      | #   log_info("Trying to find object by color:", to_str(material))
      | #   while (i < OBJECT_MAP.length()):
      | #       if (OBJECT_MAP[i].material == material):
      | #           log_info("Object model found:", to_str(OBJECT_MAP[i]))
      | #           return OBJECT_MAP[i]
      | #       end
      | #       i = i + 1
      | #   end
      | #   return OBJ_DEFAULT  # Return default pattern if not found
      | # end
      | 
      | def find_object_by_objectname(objectname):
      |     local i = 0
      |     #log_info("Trying to find object by color:", to_str(objectname))
      |     while (i < OBJECT_MAP.length()):
      |         if (OBJECT_MAP[i].obj_name == objectname):
      |             log_info("Object Model found: [" + to_str(OBJECT_MAP[i].description) + "]")
      |             return OBJECT_MAP[i]
      |         end
      |         i = i + 1
      |     end
      |     log_warning("no Object Model found for objectname:[" + to_str(objectname) + "]")
      |     return create_object()
      | end
      | 
      | def find_smallest_object():
      |     local i = 0
      |     local min_size = OBJECT_MAP[0].height
      |     #log_info("Trying to find object by color:", to_str(objectname))
      |     while (i < OBJECT_MAP.length()):
      |         if (OBJECT_MAP[i].height <= min_size and OBJECT_MAP[i].height != 0):
      |             log_info("smaller object found: [" + to_str(OBJECT_MAP[i].description) + "]")
      |             min_size = OBJECT_MAP[i].height
      |         end
      |         i = i + 1
      |     end
      |     return min_size
      | end
      | 
      | def find_gripper_config_by_objectname(objectname):
      | local i = 0
      | while (i < GRIPPER_CONFIG_MAP.length()):
      |     #log_info("gripper config:",to_str(GRIPPER_CONFIG_MAP[i]))
      |     if (GRIPPER_CONFIG_MAP[i].object == objectname):
      |         log_info("found gripper parameters [" + to_str(GRIPPER_CONFIG_MAP[i]) + "]")
      |         return GRIPPER_CONFIG_MAP[i]
      |     end
      |     i = i + 1
      | end
      | 
      | log_warning("no gripper parameters found for object type: " + to_str(objectname))
      | return create_gripper_config()
      | end
      | # Function to find a landmark by item
      | def find_landmark_by_id(lm_id):
      |     local i = 0
      |     while i < LANDMARK_MAP.length():
      |         if LANDMARK_MAP[i].lm_id == lm_id:
      |             log_info("found landmark with id(" + to_str(lm_id) + "): [" + to_str(LANDMARK_MAP[i].description) + "]")
      |             return LANDMARK_MAP[i]
      |         end
      |         i = i + 1
      |     end
      |     log_warning("landmark not found for lm_id [" + to_str(lm_id) + "]")
      |     return create_landmark()
      | end
      | # Function to find a landmark by item
      | def find_landmark_by_capture_pos(capture_pos):
      |     local i = 0
      |     while i < LANDMARK_MAP.length():
      |         if LANDMARK_MAP[i].capture_pos == capture_pos:
      |             log_info("found landmark by capture_pos [" + to_str(LANDMARK_MAP[i].description) + "]")
      |             return LANDMARK_MAP[i]
      |         end
      |         i = i + 1
      |     end
      |     log_warning("Landmark not found for capture_pos: [" + to_str(capture_pos) + "]")
      |     return create_landmark()
      | end
      | 
      | def update_landmark_by_capture_pos(capture_pos, lm_pos):
      |     local i = 0
      |     while i < LANDMARK_MAP.length():
      |         if LANDMARK_MAP[i].capture_pos == capture_pos:
      |             log_info("updated landmark from [" + to_str(LANDMARK_MAP[i].description) + "]")
      |             LANDMARK_MAP[i].actual_frame = lm_pos
      |             return True
      |         end
      |         i = i + 1
      |     end
      |     log_warning("Landmark not found for capture_pos: [" + to_str(capture_pos) + "]")
      |     return False
      | end
      | 
      | def update_landmark_by_id(lm_id,lm_pos):
      |     local i = 0
      |     while i < LANDMARK_MAP.length():
      |         if LANDMARK_MAP[i].lm_id == lm_id:
      |             log_info("updated landmark.actual_frame from [" + to_str(LANDMARK_MAP[i].description + "]"))
      |             LANDMARK_MAP[i].actual_frame = lm_pos
      |             return True
      |         end
      |         i = i + 1
      |     end
      |     log_warning("Landmark not found for lm_id " + to_str(lm_id))
      |     return False
      | end
      | 
      | def find_vision_config_by_frame(frame):
      |     local i = 0
      |     while i < VISION_CONFIG_MAP.length():
      |         if VISION_CONFIG_MAP[i].capture_pos == frame:
      |             log_info("Vision Config found: [" + to_str(VISION_CONFIG_MAP[i].description) + "]")
      |             return VISION_CONFIG_MAP[i]
      |         end
      |         i = i + 1
      |     end
      |     log_info("Vision Config not found for frame: " + to_str(frame))
      |     return create_vision_config()
      | end
      | 
      | def find_vision_config_by_itemid(id):
      |     local i = 0
      |     while i < VISION_CONFIG_MAP.length():
      |         if VISION_CONFIG_MAP[i].item_id == id:
      |             log_info("Vision Config found: [" + to_str(VISION_CONFIG_MAP[i].description) + "]")
      |             return VISION_CONFIG_MAP[i]
      |         end
      |         i = i + 1
      |     end
      |     log_info("Vision Config not found for item: " + to_str(id))
      |     return create_vision_config()
      | end
      | 
      | def find_inspect_config_by_itemid(id):
      |     local i = 0
      |     while i < INSPECT_CONFIG_MAP.length():
      |         if INSPECT_CONFIG_MAP[i].item_id == id:
      |             log_info("Inspect Config found: [" + to_str(INSPECT_CONFIG_MAP[i].description) + "]")
      |             return INSPECT_CONFIG_MAP[i]
      |         end
      |         i = i + 1
      |     end
      |     log_info("Inspect Config not found for item: " + to_str(id))
      |     return create_inspect_config()
      | end
    Script file /programs/04 Scripts/SCRIPT Device Robotiq Greifer v0.2.script
      | # ############ SCRIPT Device Robotiq Greifer ###############
      | # **********************************************************
      | # Customer          :   URG
      | # Product Name      :   uLabMobile
      | # **********************************************************
      | # Controller/Robot  :   UR5e
      | # Software          :   5.17
      | # Dependencies      :   Logs Script, Robotiq Gripper and Gripper Datastructure for args (Factory Script), URCAP Robotiq
      | # **********************************************************
      | # Author            :   D.Kreugel, P.Köhnke
      | # Copyright (c)     :   United Robotics Group Health and Food GmbH
      | #                       An der Riede 2
      | #                       28816 Stuhr
      | #                       Germany
      | # *********************************************************
      | # Description       :   Gripper Robotiq Device Interface for Robotiq E-Hand Gripper
      | # Version           :   0.2
      | # Created           :   18.07.2024
      | # Updated           :
      | # *********************************************************
      | # Modifications     :
      | #
      | # Date              :
      | # Name              :
      | # Reason            :
      | # *********************************************************
      | # TODO              :   documentation
      | 
      | # RobotiQ Gripper
      | ROBOTIQ_GRP_CLOSE = 0
      | ROBOTIQ_GRP_OPEN = 40
      | 
      | # #############FORCEMODE###############
      | ROBOTIQ_GRP_FORCE = struct(FULL=100, HALF=50, LOW=25, NONE=0)
      | 
      | # #############SPEED###################
      | ROBOTIQ_GRP_SPEED = struct(FAST=100, MEDIUM=50, SLOW=20)
      | 
      | # ############VALIDATION###############
      | ROBOTIQ_GRP_VALIDATION = struct(ON=1, OFF=0, SKIP=-1)
      | 
      | # struct(prepick=0, pick=0, place=0, force=0, speed=0, validation=0, object_type=0, description="default")
      | def gripper_robotiq_activate():
      |     return rq_activate_and_wait()
      | end
      | 
      | def gripper_robotiq_reset_and_activate():
      |     return rq_reset_and_activate()
      |     #return rq_reset()
      | end
      | 
      | def gripper_robotiq_is_activated():
      |     return rq_is_gripper_activated()
      | end
      | 
      | def gripper_robotiq_get_current_pos_mm():
      |     return rq_current_pos_mm()
      | end
      | # Function to check if the RobotiQ gripper has an object
      | def gripper_robotiq_has_object():
      |     result = rq_is_object_detected()
      |     if result == False:
      |         log_error("No object detected by the gripper")
      |     end
      |     return result
      | end
      | 
      | def gripper_robotiq_move_to_mm(mm):
      |     if(gripper_robotiq_is_activated() == False):
      |         gripper_robotiq_activate()
      |     end
      |     return rq_move_and_wait_mm(mm)
      | end
      | 
      | def gripper_robotiq_close():
      |     if(gripper_robotiq_is_activated() == False):
      |         gripper_robotiq_activate()
      |     end
      |     return rq_close_and_wait()
      | end
      | 
      | def gripper_robotiq_open():
      |     if(gripper_robotiq_is_activated() == False):
      |         gripper_robotiq_activate()
      |     end
      |     return rq_open_and_wait()
      | end
      | 
      | def gripper_robotiq_set_force(force):
      |     return rq_set_force_norm(force)
      | end
      | 
      | def gripper_robotiq_set_speed(velocity):
      |     return rq_set_speed_norm(velocity)
      | end
      | # Function to initialize the RobotiQ gripper
      | # args = struct(obj_type = object.obj_type, force = force, speed = speed, validation = validation, width = (prepick=2, pick=0, place=2))
      | def gripper_robotiq_init(args):
      |     log_info("args:"+to_str(args))
      |     gripper_robotiq_set_force(args.force)
      |     gripper_robotiq_set_speed(args.speed)
      |     if(gripper_robotiq_is_activated() == False):
      |         gripper_robotiq_activate()
      |     end
      |     log_info("Robotiq Gripper Initialized with arguments:" + to_str(args))
      |     return True
      | end
      | # Function to prepare the RobotiQ gripper for picking
      | # args = struct(obj_type = object.obj_type, force = force, speed = speed, validation = validation, width = (prepick=2, pick=0, place=2))
      | def gripper_robotiq_prepick(args):
      |     gripper_robotiq_init(args)
      | 
      |     if(args.width.prepick <= ROBOTIQ_GRP_CLOSE):
      |         rq_close_and_wait()
      |     elif(args.width.prepick >= ROBOTIQ_GRP_OPEN):
      |         rq_open_and_wait()
      |     else:
      |         rq_move_and_wait_mm(args.width.prepick)
      |     end
      | 
      |     log_info("Robotiq Gripper prepick with arguments:" + to_str(args))
      |     return True
      | end
      | 
      | # Function to place an object using the RobotiQ gripper
      | # args = struct(obj_type = object.obj_type, force = force, speed = speed, validation = validation, width = (prepick=2, pick=0, place=2))
      | def gripper_robotiq_place(args):
      |     gripper_robotiq_init(args)
      | 
      |     if(args.width.place <= ROBOTIQ_GRP_CLOSE):
      |         rq_close_and_wait()
      |     elif(args.width.place >= ROBOTIQ_GRP_OPEN):
      |         rq_open_and_wait()
      |     else:
      |         rq_move_and_wait_mm(args.width.place)
      |     end
      | 
      |     log_info("Gripper Place with arguments:"+ to_str(args))
      |     return True
      | end
      | 
      | # Function to pick an object using the RobotiQ gripper
      | # args = struct(obj_type = object.obj_type, force = force, speed = speed, validation = validation, width = (prepick=2, pick=0, place=2))
      | def gripper_robotiq_pick(args):
      |     gripper_robotiq_init(args)
      | 
      |     if(args.width.pick <= ROBOTIQ_GRP_CLOSE):
      |         rq_close_and_wait()
      |     elif(args.width.pick >= ROBOTIQ_GRP_OPEN):
      |         rq_open_and_wait()
      |     else:
      |         rq_move_and_wait_mm(args.width.pick)
      |     end
      | 
      |     log_info("Gripper Pick with arguments:" + to_str(args))
      | 
      |     if args.validation == ROBOTIQ_GRP_VALIDATION.ON:
      |         if gripper_robotiq_has_object() == False:
      |             log_error("Validation failed, no object detected")
      |             return False
      |         end
      |     end
      | 
      |     return True
      | end
      | 
      | 
      | # def gripper_robotiq_close_and_validate():
      | #     rq_close_and_wait()
      | #     if gripper_robotiq_has_object() == False:
      | #         log_error("Validation failed, no object detected")
      | #         return False
      | #     else:
      | #         return True
      | #     end
      | # end
    Script file /programs/04 Scripts/SCRIPT uLM Gripperconfig v0.6.script
      | ############# SCRIPT uLM Gripperconfig ###############
      | #*****************************************************
      | # Customer          :   URG
      | # Product Name      :   uLabMobile
      | #****************************************************
      | # Controller/Robot  :   UR5e
      | # Software          :   UR-Script
      | # Dependencies      :   physical Gripper and Datastructure from Factory for args -> Device Script and Implementations of the Functions
      | # How To            :   Assign all Functioncalls to the equivalent of the used Device Script
      | #****************************************************
      | # Author            :   D.Kreugel, P.Köhnke
      | # Copyright (c)     :   United Robotics Group Health and Food GmbH
      | #                       An der Riede 2
      | #                       28816 Stuhr
      | #                       Germany
      | #****************************************************
      | # Description       :   Defines all Gripperm related Parameters and Functions
      | # Version           :   0.6
      | # Created           :   18.07.2024
      | # Updated           :
      | #****************************************************
      | # Modifications     :   -> at the moment Gripperconfig linked to Robotiq Gripper Device Script
      | # Date              :   18.07.2017
      | # Name              :   D.Kreugel
      | # Reason            :   uLM Standard
      | #****************************************************
      | # TO DO             : Implement Activate and Reset Routine at the beginning or after an error depending on the state if an Object is gripped or not, documentation
      | 
      | 
      | 
      | # GRIPPER DEFINES
      | GRIPPER_CLOSE = ROBOTIQ_GRP_CLOSE
      | GRIPPER_OPEN = ROBOTIQ_GRP_OPEN
      | # #############FORCE###############
      | GRIPPER_FORCE = ROBOTIQ_GRP_FORCE
      | # #############SPEED###################
      | GRIPPER_SPEED = ROBOTIQ_GRP_SPEED
      | # ############VALIDATION###############
      | GRIPPER_VALIDATION = ROBOTIQ_GRP_VALIDATION
      | 
      | # takes force in %
      | def gripper_set_force(force):
      |     return gripper_robotiq_set_force(force)
      | end
      | 
      | # takes speed in %
      | def gripper_set_speed(velocity):
      |     return gripper_robotiq_set_speed(velocity)
      | end
      | 
      | def gripper_activate():
      |     return gripper_robotiq_activate()
      | end
      | 
      | def gripper_reset_and_activate():
      |     return gripper_robotiq_reset_and_activate()
      | end
      | 
      | def gripper_is_activated():
      |     return gripper_robotiq_is_activated()
      | end
      | 
      | def gripper_get_current_pos_mm():
      |     return gripper_robotiq_get_current_pos_mm()
      | end
      | 
      | def gripper_has_object():
      |     return gripper_robotiq_has_object()
      | end
      | 
      | def gripper_open():
      |     return gripper_robotiq_open()
      | end
      | 
      | def gripper_close():
      |     return gripper_robotiq_close()
      | end
      | 
      | def gripper_move_to_pos_mm(mm):
      |     return gripper_robotiq_move_to_mm(mm)
      | end
      | 
      | # args = struct(obj_type = object.obj_type, force = force, speed = speed, validation = validation, width = (prepick=2, pick=0, place=2))
      | def gripper_init(args):
      |     return gripper_robotiq_init(args)
      | end
      | 
      | # args = struct(obj_type = object.obj_type, force = force, speed = speed, validation = validation, width = (prepick=2, pick=0, place=2))
      | def gripper_prepick(args):
      |     return gripper_robotiq_prepick(args)
      | end
      | 
      | # args = struct(obj_type = object.obj_type, force = force, speed = speed, validation = validation, width = (prepick=2, pick=0, place=2))
      | def gripper_pick(args):
      |     return gripper_robotiq_pick(args)
      | end
      | 
      | # args = struct(obj_type = object.obj_type, force = force, speed = speed, validation = validation, width = (prepick=2, pick=0, place=2))
      | def gripper_place(args):
      |     return gripper_robotiq_place(args)
      | end
      | 
      | 
      | # def gripper_close_and_validate():
      | #     return gripper_robotiq_close_and_validate()
      | # end
    Script file /programs/04 Scripts/SCRIPT uLM Projectconfig 0.2.script
      | ############# SCRIPT uLM Projectconfig ###############
      | #*****************************************************
      | # Customer          :   URG
      | # Product Name      :   uLabMobile
      | #****************************************************
      | # Controller/Robot  :   UR5e
      | # Software          :   5.17
      | # Dependencies      :   Factory Script, Defines Script, relevant project knowledge about objects, patterns, items, commands, vision skills, landmarktypes and movements
      | # How To            :   Define Step by Step all Project Data by creating the objects and appending them to the assigned List, if you skip information
      | #                       the default value will be assigned -> give as many details as possible as the default values will not work in some cases
      | #****************************************************
      | # Author            :   D.Kreugel
      | # Copyright (c)     :   United Robotics Group Health and Food GmbH
      | #                       An der Riede 2
      | #                       28816 Stuhr
      | #                       Germany
      | #****************************************************
      | # Description       :   Project Related Configurations -> in the future will be configured by UGO
      | # Version           :   0.2
      | # Created           :   18.07.2024
      | # Updated           :
      | #****************************************************
      | # Modifications     :
      | # Date              :
      | # Name              :
      | # Reason            :
      | #****************************************************
      | # TO DO             :  Simplify Rack Assignment, create Enums for Choices that can be made and will be repeated in many projects, documentation
      | 
      | #
      | 
      | # Please Import DeviceScripts and Defines Script First as you may wanna use some of the Defined Variables here
      | 
      | # Define here the Objects that should be handled, add a new Object Type in the defines if necessary
      | # create_object(id=0, obj_name=0, height=0, width=0, color="default", material="default", description="default")
      | # struct(NONE=0, CC_SAMPLE=1, CC_RACK=2, COAG_SAMPLE=3, COAG_RACK=4, HEMA_SAMPLE=5, HEMA_RACK=6, INPUT_RACK=7, CF_RACK=8, ANY_SAMPLE=9, ANY_RACK=10)
      | #create_object(id=0, obj_name=0, height=0, width=0, obj_type = 0, description="default")
      | OBJECT_MAP.append(create_object(id=0, obj_name=Objects.NONE, obj_type=ObjectType.NONE, height=0, width=0, description="None Object"))
      | OBJECT_MAP.append(create_object(id=1, obj_name=Objects.CC_SAMPLE, obj_type=ObjectType.SAMPLE, height=108, width=15, description="BD Li-Heparin"))
      | OBJECT_MAP.append(create_object(id=2, obj_name=Objects.HEMA_SAMPLE, obj_type=ObjectType.SAMPLE, height=81, width=13, description="BD EDTA"))
      | OBJECT_MAP.append(create_object(id=3, obj_name=Objects.CC_SAMPLE, obj_type=ObjectType.SAMPLE, height=108, width=15, description="BD Li-Heparin"))
      | OBJECT_MAP.append(create_object(id=4, obj_name=Objects.HEMA_SAMPLE, obj_type=ObjectType.SAMPLE, height=81, width=13, description="Sarstedt EDTA"))
      | OBJECT_MAP.append(create_object(id=5, obj_name=Objects.CC_SAMPLE, obj_type=ObjectType.SAMPLE, height=110, width=15, description="Sarstedt Serum-Gel"))
      | OBJECT_MAP.append(create_object(id=6, obj_name=Objects.ANY_SAMPLE, obj_type=ObjectType.SAMPLE, height=110, width=15, description="Any Sample"))
      | OBJECT_MAP.append(create_object(id=7, obj_name=Objects.ANY_RACK, height=150, width=120, description="Any Rack"))
      | OBJECT_MAP.append(create_object(id=8, obj_name=Objects.CF_RACK, height=110, width=15, description="Centrifuge Rack"))
      | OBJECT_MAP.append(create_object(id=12, obj_name=Objects.COBAS_RACK, height=OBJECT_REFERENCE_HEIGHT, width=20, description="Cobas Rack"))
      | OBJECT_MAP.append(create_object(id=9, obj_name=Objects.TARA_SAMPLE, obj_type=ObjectType.SAMPLE, height=110, width=15, description="Tara Sample"))
      | OBJECT_MAP.append(create_object(id=10, obj_name=Objects.BUTTON, obj_type=ObjectType.BUTTON, height=0, width=0, description="Button"))
      | OBJECT_MAP.append(create_object(id=11, obj_name=Objects.XN550_DRAWER, height=OBJECT_REFERENCE_HEIGHT, width=25, description="XN550 Drawer"))
      | 
      | #create_sample(obj_id=0, diameter=0, color="", material="", description="")
      | SAMPLES = make_list(0,create_sample(),MAX_ITEM_OBJ)
      | SAMPLES.append(create_sample(obj_id=1, cap_diameter=17.4, raw_diameter=15.3, color="darkgreen", material="88", description="BD Li-Heparin -> decapped in Cobas"))
      | SAMPLES.append(create_sample(obj_id=1, cap_diameter=17.4, raw_diameter=15.3, color="darkgreen", material="80", description="BD Li-Heparin -> decapped in Cobas"))
      | SAMPLES.append(create_sample(obj_id=1, cap_diameter=17.4, raw_diameter=15.3, color="darkgreen", material="93", description="BD Li-Heparin -> decapped in archive"))
      | SAMPLES.append(create_sample(obj_id=2, cap_diameter=15.5, raw_diameter=12.3, color="violet", material="82", description="BD EDTA -> Sysmex ->Archive"))
      | SAMPLES.append(create_sample(obj_id=2, cap_diameter=15.5, raw_diameter=12.3, color="violet", material="91", description="BD EDTA ->Archive"))
      | SAMPLES.append(create_sample(obj_id=2, cap_diameter=15.5, raw_diameter=12.3, color="violet", material="96", description="BD EDTA ->Archive"))
      | SAMPLES.append(create_sample(obj_id=3, cap_diameter=17.4, raw_diameter=15.3, color="lightgreen", material="88", description="BD Li-Heparin -> decapped in Cobas"))
      | SAMPLES.append(create_sample(obj_id=3, cap_diameter=17.4, raw_diameter=15.3, color="lightgreen", material="93", description="BD Li-Heparin -> decapped in Archive"))
      | SAMPLES.append(create_sample(obj_id=3, cap_diameter=17.4, raw_diameter=15.3, color="lightgreen", material="97", description="BD Li-Heparin -> decapped in Archive"))
      | SAMPLES.append(create_sample(obj_id=4, cap_diameter=15.6, raw_diameter=12.3, color="red", material="82", description="BD EDTA -> Sysmex ->Archive"))
      | SAMPLES.append(create_sample(obj_id=4, cap_diameter=15.6, raw_diameter=12.3, color="red", material="91", description="BD EDTA -> Archive"))
      | SAMPLES.append(create_sample(obj_id=4, cap_diameter=15.6, raw_diameter=12.3, color="red", material="96", description="BD EDTA -> Archive"))
      | SAMPLES.append(create_sample(obj_id=5, cap_diameter=17.4, raw_diameter=15.3, color="brown", material="80", description="Sarstedt Serum-Gel -> decapped in Cobas"))
      | SAMPLES.append(create_sample(obj_id=5, cap_diameter=17.4, raw_diameter=15.3, color="brown", material="93", description="Sarstedt Serum-Gel -> decapped in Archive"))
      | 
      | # Gripper Configurations depending on the Object Type , add new force and speed in the Defines if necessary
      | # create_gripper_config(gripper_offset=struct(prepick=2, pick=0, place=2), force=0, speed=0, validation=0, object=create_object())
      | GRIPPER_CONFIG_MAP.append(create_gripper_config(gripper_offset=struct(prepick=2, pick=0, place=2), force=GRIPPER_FORCE.HALF, speed=GRIPPER_SPEED.MEDIUM, validation=GRIPPER_VALIDATION.ON, object=find_object_by_objectname(Objects.ANY_SAMPLE)))
      | GRIPPER_CONFIG_MAP.append(create_gripper_config(gripper_offset=struct(prepick=2, pick=0, place=2), force=GRIPPER_FORCE.FULL, speed=GRIPPER_SPEED.MEDIUM, validation=GRIPPER_VALIDATION.ON, object=find_object_by_objectname(Objects.ANY_RACK)))
      | GRIPPER_CONFIG_MAP.append(create_gripper_config(gripper_offset=struct(prepick=2, pick=0, place=2), force=GRIPPER_FORCE.HALF, speed=GRIPPER_SPEED.MEDIUM, validation=GRIPPER_VALIDATION.ON, object=find_object_by_objectname(Objects.CC_SAMPLE)))
      | GRIPPER_CONFIG_MAP.append(create_gripper_config(gripper_offset=struct(prepick=3, pick=0, place=3), force=GRIPPER_FORCE.HALF, speed=GRIPPER_SPEED.MEDIUM, validation=GRIPPER_VALIDATION.ON, object=find_object_by_objectname(Objects.HEMA_SAMPLE)))
      | GRIPPER_CONFIG_MAP.append(create_gripper_config(gripper_offset=struct(prepick=4, pick=0, place=4), force=GRIPPER_FORCE.HALF, speed=GRIPPER_SPEED.MEDIUM, validation=GRIPPER_VALIDATION.OFF, object=find_object_by_objectname(Objects.TARA_SAMPLE)))
      | GRIPPER_CONFIG_MAP.append(create_gripper_config(gripper_offset=struct(prepick=2, pick=0, place=2), force=GRIPPER_FORCE.FULL, speed=GRIPPER_SPEED.MEDIUM, validation=GRIPPER_VALIDATION.ON, object=find_object_by_objectname(Objects.CF_RACK)))
      | GRIPPER_CONFIG_MAP.append(create_gripper_config(gripper_offset=struct(prepick=2, pick=0, place=2), force=GRIPPER_FORCE.FULL, speed=GRIPPER_SPEED.MEDIUM, validation=GRIPPER_VALIDATION.ON, object=find_object_by_objectname(Objects.COBAS_RACK)))
      | GRIPPER_CONFIG_MAP.append(create_gripper_config(gripper_offset=struct(prepick=0, pick=0, place=0), force=GRIPPER_FORCE.HALF, speed=GRIPPER_SPEED.MEDIUM, validation=GRIPPER_VALIDATION.OFF, object=find_object_by_objectname(Objects.NONE)))
      | GRIPPER_CONFIG_MAP.append(create_gripper_config(gripper_offset=struct(prepick=0, pick=0, place=0), force=GRIPPER_FORCE.HALF, speed=GRIPPER_SPEED.MEDIUM, validation=GRIPPER_VALIDATION.OFF, object=find_object_by_objectname(Objects.BUTTON)))
      | GRIPPER_CONFIG_MAP.append(create_gripper_config(gripper_offset=struct(prepick=5, pick=25, place=5), force=GRIPPER_FORCE.HALF, speed=GRIPPER_SPEED.MEDIUM, validation=GRIPPER_VALIDATION.OFF, object=find_object_by_objectname(Objects.XN550_DRAWER)))
      | # create Patterns like Racks or Magazines
      | # easy if you define x and y regarding to the base coordinate system  if not you have to deal with transpose and or invert
      | # create_pattern(id=0, pattern_width=[0, 0], pattern_size=[0, 0], blocked=[-1, -1], obj_name=0, direction="X", transpose=False, invert=False, description="default")
      | # Objectss: NONE=0, CC_SAMPLE=1, CC_RACK=2, COAG_SAMPLE=3, COAG_RACK=4, HEMA_SAMPLE=5, HEMA_RACK=6, INPUT_RACK=7, CENTRIFUGE_RACK=8, ANY_SAMPLE=9, ANY_RACK=10
      | # ITEM_MODEL_MAP.append(create_pattern(id=0, pattern_width=[0, 0], pattern_size=[0, 0], blocked=[-1, -1, -1],  direction="X", transpose=False, invert=False, description="default"))
      | # ITEM_MODEL_MAP.append(create_pattern(id=1, pattern_width=[0.06, 0], pattern_size=[3, 1],  direction="X", description="Tara"))
      | # ITEM_MODEL_MAP.append(create_pattern(id=2, pattern_width=[0.183, 0.082], pattern_size=[10, 5], description="Sarstedt 50 D17 Rack"))
      | # ITEM_MODEL_MAP.append(create_pattern(id=3, pattern_width=[0.153, 0.067], pattern_size=[10, 5], description="Sarstedt 50 D13 Rack"))
      | # ITEM_MODEL_MAP.append(create_pattern(id=4, pattern_width=[0.06, 0.06], pattern_size=[3, 3], blocked=[5, -1, -1], description="Hettich Centrifuge Rack"))
      | # ITEM_MODEL_MAP.append(create_pattern(id=5, pattern_width=[0.093, 0.093], pattern_size=[2, 2],  description="Hettich Centrifuge Rack Magazin"))
      | # ITEM_MODEL_MAP.append(create_pattern(id=6, pattern_width=[0.08, 0.05], pattern_size=[5, 2], description="Sysmex XN 550 Rack"))
      | # ITEM_MODEL_MAP.append(create_pattern(id=7, pattern_width=[0.175, 0.078], pattern_size=[8, 4], description="URG Rack 40 D17"))
      | # ITEM_MODEL_MAP.append(create_pattern(id=8, pattern_width=[0.092, 0], pattern_size=[5, 1], description="Cobas Rack"))
      | # ITEM_MODEL_MAP.append(create_pattern(id=9, pattern_width=[0.245, 0.123], pattern_size=[3, 5], blocked=[9,11,12], description="Cobas Rack Magazin"))
      | # ITEM_MODEL_MAP.append(create_pattern(id=10, pattern_width=[0.237, 0.095], pattern_size=[11, 5], description="Atellica Rack 5x11"))
      | # ITEM_MODEL_MAP.append(create_pattern(id=11, pattern_width=[0.237, 0.095], pattern_size=[2, 2], description="Sensors LM"))
      | # ITEM_MODEL_MAP.append(create_pattern(id=12, pattern_width=[0.18, 0], pattern_size=[10, 1], description="Sysmex CS2500 Rack"))
      | # ITEM_MODEL_MAP.append(create_pattern(id=13, pattern_width=[0.310, 0.075], pattern_size=[13, 4], description="URG RACK 52 - Special Input"))
      | # ITEM_MODEL_MAP.append(create_pattern(id=14, pattern_width=[0.075, 0.075], pattern_size=[4, 6], description="URG RACK 24 - Special NoK"))
      | # ITEM_MODEL_MAP.append(create_pattern(id=15, pattern_width=[0.120, 0], pattern_size=[2, 1], description="XN550 Drawer"))
      | 
      | ITEM_MODEL_MAP.append(create_pattern(id=0, name="NONE", pattern_width=[0, 0], pattern_size=[0, 0], blocked=[-1, -1, -1],  direction="X", transpose=False, invert=False, description="default"))
      | ITEM_MODEL_MAP.append(create_pattern(id=1, name="TARA", pattern_width=[0.06, 0], pattern_size=[3, 1],  direction="X", description="Tara"))
      | ITEM_MODEL_MAP.append(create_pattern(id=4, name="CENTRIFUGE", pattern_width=[0.06, 0.06], pattern_size=[3, 3], blocked=[5, -1, -1], description="Hettich Centrifuge Rack"))
      | ITEM_MODEL_MAP.append(create_pattern(id=5, name="CENTRIFUGE_MAGAZINE", pattern_width=[0.093, 0.093], pattern_size=[2, 2],  description="Hettich Centrifuge Rack Magazin"))
      | ITEM_MODEL_MAP.append(create_pattern(id=6, name="SYSMEX_XN550", pattern_width=[0.08, 0.05], pattern_size=[5, 2], description="Sysmex XN 550 Rack"))
      | ITEM_MODEL_MAP.append(create_pattern(id=8, name="COBAS", pattern_width=[0.092, 0], pattern_size=[5, 1], description="Cobas Rack"))
      | ITEM_MODEL_MAP.append(create_pattern(id=9, name="COBAS_MAGAZINE", pattern_width=[0.245, 0.123], pattern_size=[3, 5], blocked=[9,11,12], description="Cobas Rack Magazin"))
      | ITEM_MODEL_MAP.append(create_pattern(id=13, name="INPUT", pattern_width=[0.310, 0.075], pattern_size=[13, 4], description="URG RACK 52 - Special Input"))
      | ITEM_MODEL_MAP.append(create_pattern(id=14, name="NOK", pattern_width=[0.075, 0.075], pattern_size=[4, 6], description="URG RACK 24 - Special NoK"))
      | ITEM_MODEL_MAP.append(create_pattern(id=15, name="DRAWER_XN550", pattern_width=[0.120, 0], pattern_size=[2, 1], description="XN550 Drawer"))
      | ITEM_MODEL_MAP.append(create_pattern(id=7, name="ARCHIVE", pattern_width=[0.175, 0.078], pattern_size=[8, 4], description="URG Rack 40 D17"))
      | 
      | 
      | 
      | 
      | 
      | 
      | # add a "skill" to the robots skillset the control system will send a string with the ls_item and action and here we will look if we have a matching skill to execute
      | # the item_modell defines the patterns which have to be used by the robot on multiple racks and or multiple samples in a rackpattern
      | # inner pattern is always dependung on the object that has to be moved and the outer pattern is the pattern for the containers where the objects are stored in.
      | # if racks have to be handled it is also an inner pattern cause the object to handle is the rack itself
      | # create_item(id=0, ls_item="default", frame=p[0,0,0,0,0,0], actionlist=create_action_list([]), item_model=create_item_model(), lm_id=0, description="default")
      | # create_item_model(inner=create_pattern(), outer=create_pattern(), description="default")
      | # ITEM_MAP.append(create_item(id=1, ls_item="Home", frame=F1_uLM_Home, actionlist=[ActionManipulator.MOVE_TO], description="uLM Move To Home"))
      | # ITEM_MAP.append(create_item(id=2, ls_item="InputStation", frame=F2_uLM_Input, actionlist=[ActionManipulator.PICK, ActionManipulator.PLACE], item_model=create_item_model(inner=Patterns.INPUT), description="uLM Pick and Place samples from Input"))
      | # ITEM_MAP.append(create_item(id=3, ls_item="InputCapture", frame=F3_Cap_Input, actionlist=[ActionCamera.INSPECT, ActionManipulator.MOVE_TO], description="uLM Inspect samples from Input and Move To Capture Position"))
      | # ITEM_MAP.append(create_item(id=4, ls_item="Bin", frame=F4_uLM_Bin, actionlist=[ActionManipulator.PLACE], description="uLM Place Cap to Bin"))
      | # ITEM_MAP.append(create_item(id=5, ls_item="StationaryGripper", frame=F5_uLM_Gripper, actionlist=[ActionManipulator.PICK, ActionManipulator.PLACE, ActionManipulator.DECAP, ActionManipulator.MOVE_TO, ActionManipulator.GRASP, ActionManipulator.RELEASE], description=" uLM stationary gripper"))
      | # ITEM_MAP.append(create_item(id=6, ls_item="CobasRack", frame=F6_uLM_Cobas_R, actionlist=[ActionManipulator.PICK, ActionManipulator.PLACE], item_model=create_item_model(outer=Patterns.COBAS_MAGAZINE), description="uLM Cobas Racks Pick and Place"))
      | # ITEM_MAP.append(create_item(id=7, ls_item="CobasMagazine", frame=F7_uLM_Coba_Mag, actionlist=[ActionManipulator.PICK, ActionManipulator.PLACE], item_model=create_item_model(inner=Patterns.COBAS, outer=Patterns.COBAS_MAGAZINE), description="uLM Cobas Magazine Samples Pick and Place"))
      | # ITEM_MAP.append(create_item(id=8, ls_item="DetectCobasRacks", frame=F8_Cap_Cobas_LM, actionlist=[ActionCamera.DETECT_OBJECTS, ActionManipulator.MOVE_TO], lm_id=2, description="uLM Cobas Rack Detection and Move To Capture"))
      | # ITEM_MAP.append(create_item(id=9, ls_item="TaraMagazine", frame=F9_uLM_Tara, actionlist=[ActionManipulator.PICK, ActionManipulator.PLACE], item_model=create_item_model(inner=Patterns.TARA), description="uLM Centrifuge Tara Pick and Place"))
      | # ITEM_MAP.append(create_item(id=10, ls_item="CentrifugeCapture", frame=F10_Cap_CF, actionlist=[ActionManipulator.MOVE_TO, ActionCamera.DETECT], lm_id=1, description="Centrifuge Device Move to Capture Pos and Detect Landmarks"))
      | # ITEM_MAP.append(create_item(id=11, ls_item="Centrifuge", frame=F11_CF_PiPl, actionlist=[ActionManipulator.PICK, ActionManipulator.PLACE], description="Centrifuge Device Rack Pick and Place"))
      | # ITEM_MAP.append(create_item(id=12, ls_item="CentrifugeMagazine", frame=F12_uLM_CF_Mag, actionlist=[ActionManipulator.PICK, ActionManipulator.PLACE], item_model=create_item_model(inner=Patterns.CENTRIFUGE, outer=Patterns.CENTRIFUGE_MAGAZINE), description=" uLM Centrifuge Magazin Pick and Place"))
      | # ITEM_MAP.append(create_item(id=13, ls_item="CentrifugeRack", frame=F13_uLM_CF_R, actionlist=[ActionManipulator.PICK, ActionManipulator.PLACE], item_model=create_item_model(outer=Patterns.CENTRIFUGE_MAGAZINE), description="uLM Centrifuge Magazin Pick and Place Racks"))
      | # ITEM_MAP.append(create_item(id=14, ls_item="DailyArchive", frame=F14_uLM_Archive, actionlist=[ActionManipulator.PICK, ActionManipulator.PLACE], item_model=create_item_model(inner=Patterns.ARCHIVE), description="uLM Pick and Place samples from Archive Rack"))
      | # ITEM_MAP.append(create_item(id=15, ls_item="NokRack", frame=F15_uLM_Nok, actionlist=[ActionManipulator.PICK, ActionManipulator.PLACE], item_model=create_item_model(inner=Patterns.NOK), description="uLM Pick and Place samples from Nok Rack"))
      | # ITEM_MAP.append(create_item(id=16, ls_item="CobasInput", frame=F16_Cobas_Input, actionlist=[ActionManipulator.PLACE], description="uLM Place Cobasrack in Cobas Device"))
      | # ITEM_MAP.append(create_item(id=17, ls_item="CobasInputCapture", frame=F17_Cobas_Cap, actionlist=[ActionCamera.DETECT, ActionManipulator.MOVE_TO], lm_id=3, description="uLM Place Cobasrack in Cobas Device"))
      | # ITEM_MAP.append(create_item(id=18, ls_item="XN550Input", frame=F18_XN550_Input, actionlist=[ActionManipulator.PICK, ActionManipulator.PLACE], item_model=create_item_model(inner=Patterns.SYSMEX_XN550, outer=Patterns.DRAWER_XN550), lm_id=4, description="uLM Pick and Place Samples in or out of XN550 Racks"))
      | # ITEM_MAP.append(create_item(id=19, ls_item="XN550Capture", frame=F19_XN550_Cap, actionlist=[ActionCamera.DETECT, ActionManipulator.MOVE_TO], lm_id=4, description="uLM Move To and Capture LM XN550"))
      | # ITEM_MAP.append(create_item(id=20, ls_item="XN550Drawer", frame=F20_XN550_Draw, actionlist=[ActionManipulator.DRAWER_OPEN, ActionManipulator.DRAWER_CLOSE], item_model=create_item_model(inner=Patterns.DRAWER_XN550), lm_id=4, description="uLM Open and close Drawer XN550"))
      | # ITEM_MAP.append(create_item(id=21, ls_item="XN550Button", frame=F21_XN550_Btn, actionlist=[ActionManipulator.PUSH], lm_id=4, description="uLM Push XN550 Button"))
      | # ITEM_MAP.append(create_item(id=22, ls_item="AMR", frame=p[0,0,0,0,0,0], actionlist=[ActionAMR.READ, ActionAMR.LOAD_MISSION, ActionAMR.START_MISSION, ActionAMR.NAVIGATE, ActionAMR.ACKNOWLEDGE], description="all AMR actions"))
      | 
      | 
      | 
      | # ITEM_MAP.append(create_item(id=31, ls_item="TestLM", frame=TestLM, actionlist=[ActionManipulator.PICK, ActionManipulator.PLACE], item_model=create_item_model(inner=Rack.SYSMEX_CS2500), lm_id=5, description="LM Test"))
      | # Fills the Vision Config List with Projectrelated Data
      | # workspaceid and skillid are highly robominds related so probably will not stay like this in the future
      | # sample detection: dx and dy are used to calculate the positions in a rack and given by the offset which will be applied in order to assign the sample to a place in the rack
      | # create_vision_config(workspace_id="", skill_id="", item_id=-1, capture_pos=p[0,0,0,0,0,0], dx=0, dy=0, target_origin=p[0,0,0,0,0,0], selector="default", description="default")
      | # VISION_CONFIG_MAP.append(create_vision_config(workspace_id="96017791-f581-4e9e-93da-6951695fccc8", skill_id="8885cfe1-6784-4293-bd26-52ebdc67bf95", capture_pos=F10_Cap_CF, target_origin=p[0,0,0,0,0,0], item_id=11, description="LM Detect CF"))
      | # VISION_CONFIG_MAP.append(create_vision_config(workspace_id="96017791-f581-4e9e-93da-6951695fccc8", skill_id="8885cfe1-6784-4293-bd26-52ebdc67bf95", capture_pos=F8_Cap_Cobas_LM, target_origin=p[0,0,0,0,0,0], item_id=8, description="LM Detect Cobas Racks"))
      | # VISION_CONFIG_MAP.append(create_vision_config(workspace_id="8f0ad01c-dc36-4fdd-b295-0b6b4a38b89a", skill_id="afdc9e13-ea83-40d6-a805-bb041453d2e5", capture_pos=F3_Cap_Input, target_origin=F2_uLM_Input, item_id=3, description="Lab Solution Input Capture"))
      | # VISION_CONFIG_MAP.append(create_vision_config(workspace_id="96017791-f581-4e9e-93da-6951695fccc8", skill_id="8885cfe1-6784-4293-bd26-52ebdc67bf95", capture_pos=F19_XN550_Cap, target_origin=F18_XN550_Input, item_id=18, description="Input XN550"))
      | # VISION_CONFIG_MAP.append(create_vision_config(workspace_id="96017791-f581-4e9e-93da-6951695fccc8", skill_id="8885cfe1-6784-4293-bd26-52ebdc67bf95", capture_pos=F19_XN550_Cap, target_origin=POS_Z, item_id=19, description="LM Detect XN550F"))
      | # VISION_CONFIG_MAP.append(create_vision_config(workspace_id="96017791-f581-4e9e-93da-6951695fccc8", skill_id="8885cfe1-6784-4293-bd26-52ebdc67bf95", capture_pos=F10_Cap_CF, target_origin=POS_Z, item_id=10, description="LM Detect CF"))
      | # VISION_CONFIG_MAP.append(create_vision_config(workspace_id="96017791-f581-4e9e-93da-6951695fccc8", skill_id="8885cfe1-6784-4293-bd26-52ebdc67bf95", capture_pos=F19_XN550_Cap, target_origin=F20_XN550_Draw, item_id=20, description="Drawer XN550"))
      | # VISION_CONFIG_MAP.append(create_vision_config(workspace_id="96017791-f581-4e9e-93da-6951695fccc8", skill_id="8885cfe1-6784-4293-bd26-52ebdc67bf95", capture_pos=F19_XN550_Cap, target_origin=F21_XN550_Btn, item_id=21, description="Button XN550"))
      | # VISION_CONFIG_MAP.append(create_vision_config(workspace_id="96017791-f581-4e9e-93da-6951695fccc8", skill_id="8885cfe1-6784-4293-bd26-52ebdc67bf95", capture_pos=TestLMCap, target_origin=p[0,0,0,0,0,0], item_id=30, description="Button XN550"))
      | # VISION_CONFIG_MAP.append(create_vision_config(workspace_id="96017791-f581-4e9e-93da-6951695fccc8", skill_id="8885cfe1-6784-4293-bd26-52ebdc67bf95", capture_pos=TestLMCap, target_origin=TestLM, item_id=31, description="Button XN550"))
      | 
      | # VISION_CONFIG_MAP.append(create_vision_config(workspace_id="96017791-f581-4e9e-93da-6951695fccc8", skill_id="8885cfe1-6784-4293-bd26-52ebdc67bf95", target_origin=p[0,0,0,0,0,0], item_id=11, description="LM Detect CF"))
      | # VISION_CONFIG_MAP.append(create_vision_config(workspace_id="96017791-f581-4e9e-93da-6951695fccc8", skill_id="8885cfe1-6784-4293-bd26-52ebdc67bf95", target_origin=p[0,0,0,0,0,0], item_id=8, description="LM Detect Cobas Racks"))
      | # VISION_CONFIG_MAP.append(create_vision_config(workspace_id="8f0ad01c-dc36-4fdd-b295-0b6b4a38b89a", skill_id="afdc9e13-ea83-40d6-a805-bb041453d2e5", target_origin=F2_uLM_Input, item_id=3, description="Lab Solution Input Capture"))
      | # VISION_CONFIG_MAP.append(create_vision_config(workspace_id="96017791-f581-4e9e-93da-6951695fccc8", skill_id="8885cfe1-6784-4293-bd26-52ebdc67bf95", target_origin=F18_XN550_Input, item_id=18, description="Input XN550"))
      | # VISION_CONFIG_MAP.append(create_vision_config(workspace_id="96017791-f581-4e9e-93da-6951695fccc8", skill_id="8885cfe1-6784-4293-bd26-52ebdc67bf95", target_origin=POS_Z, item_id=19, description="LM Detect XN550F"))
      | # VISION_CONFIG_MAP.append(create_vision_config(workspace_id="96017791-f581-4e9e-93da-6951695fccc8", skill_id="8885cfe1-6784-4293-bd26-52ebdc67bf95", target_origin=POS_Z, item_id=10, description="LM Detect CF"))
      | # VISION_CONFIG_MAP.append(create_vision_config(workspace_id="96017791-f581-4e9e-93da-6951695fccc8", skill_id="8885cfe1-6784-4293-bd26-52ebdc67bf95", target_origin=F20_XN550_Draw, item_id=20, description="Drawer XN550"))
      | # VISION_CONFIG_MAP.append(create_vision_config(workspace_id="96017791-f581-4e9e-93da-6951695fccc8", skill_id="8885cfe1-6784-4293-bd26-52ebdc67bf95", target_origin=F21_XN550_Btn, item_id=21, description="Button XN550"))
      | # VISION_CONFIG_MAP.append(create_vision_config(workspace_id="96017791-f581-4e9e-93da-6951695fccc8", skill_id="8885cfe1-6784-4293-bd26-52ebdc67bf95", target_origin=p[0,0,0,0,0,0], item_id=30, description="Button XN550"))
      | # VISION_CONFIG_MAP.append(create_vision_config(workspace_id="96017791-f581-4e9e-93da-6951695fccc8", skill_id="8885cfe1-6784-4293-bd26-52ebdc67bf95", target_origin=TestLM, item_id=31, description="Button XN550"))
      | 
      | # local inputrack = find_pattern_by_name("INPUT")
      | # INSPECT_CONFIG_MAP.append(create_inspect_config(item_id=3, dx=inputrack.pattern_width[0]/(inputrack.pattern_size[0]-1), dy=inputrack.pattern_width[1]/(inputrack.pattern_size[1]-1), rack_size=inputrack.pattern_size , description="Input Capture"))
      | # # Fills the Landmark List with Projectrelated Data
      | # # create_landmark(lm_id=0, marker_id=-1, marker_size=0.1, marker_type="aruco_7x7", capture_pos=p[0,0,0,0,0,0], init_frame=p[0,0,0,0,0,0], search_offset=[0,0,0], actual_frame=p[0,0,0,0,0,0], description="")
      | # LANDMARK_MAP.append(create_landmark(lm_id=1, marker_id=3, marker_size=0.1, marker_type="aruco_7x7", capture_pos = F10_Cap_CF, init_frame=p[-0.617789, -0.065471, 0.07918, 0.020983, -0.012695, 1.512066], search_offset=[0.15, 0.15, 0.1], actual_frame=p[-0.617789, -0.065471, 0.07918, 0.020983, -0.012695, 1.512066], description="LM CF Lid"))
      | # LANDMARK_MAP.append(create_landmark(lm_id=2, marker_id=-1, marker_size=0.0085, marker_type="aruco_4x4", capture_pos = F8_Cap_Cobas_LM, init_frame=p[0,0,0,0,0,0], search_offset=[0.15, 0.15, 0.1], actual_frame=POS_Z, description="LM Cobas Rack Detection"))
      | # LANDMARK_MAP.append(create_landmark(lm_id=3, marker_id=0, marker_size=0.1, marker_type="aruco_7x7", capture_pos = F17_Cobas_Cap, init_frame=p[-0.667,-0.194,0.100,0,0,0], search_offset=[0.15, 0.15, 0.1], actual_frame=POS_Z, description="LM Cobas Cap"))
      | # LANDMARK_MAP.append(create_landmark(lm_id=4, marker_id=4, marker_size=0.1, marker_type="aruco_7x7", capture_pos = F19_XN550_Cap, init_frame=p[0.124,-0.976,0.355,-0.008,0.025,3.131], search_offset=[0.15, 0.15, 0.1], actual_frame=p[0,0,0,0,0,0], description="LM XN550 Cap"))
      | # LANDMARK_MAP.append(create_landmark(lm_id=5, marker_id=0, marker_size=0.1, marker_type="aruco_7x7", capture_pos = TestLMCap, init_frame=p[-0.49,-0.144,0.092,0,-0.008,0.001], search_offset=[0.15, 0.15, 0.1], actual_frame=POS_Z, description="LM Test"))
      | # # Configuration of all movement related parameters
      | # # create_movement(id=0, hh_approach=POS_Z, h_approach=POS_Z, approach=POS_Z, h_target=POS_Z, target=POS_Z, retract=POS_Z, h_retract=POS_Z, hh_retract=POS_Z, h_frame=POS_Z, frame=POS_Z, speed=1, acceleration=1, description="default")
      | # MOVEMENT_MAP.append(create_movement(description="TestLMCap", frame=TestLMCap, actionlist=[ActionManipulator.MOVE_TO]))
      | # MOVEMENT_MAP.append(create_movement(description="TestLM", frame=TestLM, actionlist=[ActionManipulator.PICK,ActionManipulator.PLACE],
      | #         approach=p[0,0,0.1,0,0,0],
      | #         retract=p[0,0,0.1,0,0,0]))
      | # MOVEMENT_MAP.append(create_movement(description="Home - MOVE_TO", frame=F1_uLM_Home, actionlist=[ActionManipulator.MOVE_TO]))
      | # MOVEMENT_MAP.append(create_movement(description="Input - PICK&PLACE", frame=F2_uLM_Input, actionlist=[ActionManipulator.PICK,ActionManipulator.PLACE],
      | #         approach=p[0,0,0.1,0,0,0],
      | #         retract=p[0,0,0.1,0,0,0]))
      | # MOVEMENT_MAP.append(create_movement(description="Capture Input - MOVE_TO", frame=F3_Cap_Input, actionlist=[ActionManipulator.MOVE_TO]))
      | # MOVEMENT_MAP.append(create_movement(description="BIN - PLACE", frame=F4_uLM_Bin, actionlist=[ActionManipulator.PLACE],
      | #         approach=p[0,0,0.1,0,0,0],
      | #         retract=p[0,0,0.1,0,0,0]))
      | # MOVEMENT_MAP.append(create_movement(description="Gripper - Move To", frame=F5_uLM_Gripper, actionlist=[ActionManipulator.MOVE_TO],
      | #         approach=p[0,0,0.1,0,0,0]))
      | # MOVEMENT_MAP.append(create_movement(description="Gripper - Pick", frame=F5_uLM_Gripper, actionlist=[ActionManipulator.PICK],
      | #         retract=p[0,0,0.1,0,0,0]))
      | # MOVEMENT_MAP.append(create_movement(description="Gripper - Place", frame=F5_uLM_Gripper, actionlist=[ActionManipulator.PLACE],
      | #         approach=p[0,0,0.1,0,0,0]))
      | # MOVEMENT_MAP.append(create_movement(description="CobasRack Pick & Place", frame=F6_uLM_Cobas_R, actionlist=[ActionManipulator.PICK,ActionManipulator.PLACE],
      | #         approach=p[0,0,0.1,0,0,0],
      | #         target=p[0,0,0,0,0,d2r(90)],
      | #         retract=p[0,0,0.1,0,0,0]))
      | # MOVEMENT_MAP.append(create_movement(description="CobasMagazine Pick & Place", frame=F7_uLM_Coba_Mag, actionlist=[ActionManipulator.PICK,ActionManipulator.PLACE],
      | #         approach=p[0,0,0.1,0,0,0],
      | #         target=p[0,0,0,0,0,-d2r(90)],
      | #         retract=p[0,0,0.1,0,0,0]))
      | # MOVEMENT_MAP.append(create_movement(description="Capture Position Cobas Landmarks", frame=F8_Cap_Cobas_LM, actionlist=[ActionManipulator.MOVE_TO]))
      | # MOVEMENT_MAP.append(create_movement(description="TaraMagazine - PICK & PLACE", frame=F9_uLM_Tara, actionlist=[ActionManipulator.PICK,ActionManipulator.PLACE],
      | #         approach=p[0,0,0.13,0,0,0],
      | #         target=p[0,0,0,0,0,-d2r(90)],
      | #         retract=p[0,0,0.13,0,0,0]))
      | # MOVEMENT_MAP.append(create_movement(description="Capture Position - Centrifuge LM", frame=F10_Cap_CF,actionlist=[ActionManipulator.MOVE_TO]))
      | # MOVEMENT_MAP.append(create_movement(description="Pick and Place Racks - Centrifuge Lid", frame=F11_CF_PiPl, actionlist=[ActionManipulator.PICK,ActionManipulator.PLACE],
      | #         approach=p[0,0,0.3,0,0,0],
      | #         retract=p[0,0,0.3,0,0,0]))
      | # MOVEMENT_MAP.append(create_movement(description="Pick and Place Samples - Centrifuge on uLM", frame=F12_uLM_CF_Mag, actionlist=[ActionManipulator.PICK,ActionManipulator.PLACE],
      | #         approach=p[0,0,0.13,0,0,0],
      | #         retract=p[0,0,0.13,0,0,0]
      | #         ))
      | # MOVEMENT_MAP.append(create_movement(description="Pick and Place Racks - Centrifuge on uLM", frame=F13_uLM_CF_R, actionlist=[ActionManipulator.PICK,ActionManipulator.PLACE],
      | #         approach=p[0,0,0.15,0,0,0],
      | #         retract=p[0,0,0.15,0,0,0]
      | #         ))
      | 
      | # MOVEMENT_MAP.append(create_movement(description="Pick and Place Samples XN550 Racks in Device", frame=F18_XN550_Input, actionlist=[ActionManipulator.PICK,ActionManipulator.PLACE],
      | #         approach=p[0,0,0.1,0,0,0],
      | #         target = p[0,0,0,0,0,d2r(90)],
      | #         retract=p[0,0,0.1,0,0,0]
      | #         ))
      | # MOVEMENT_MAP.append(create_movement(description="Capture LM XN550", frame=F19_XN550_Cap, actionlist=[ActionManipulator.MOVE_TO]))
      | # MOVEMENT_MAP.append(create_movement(description="Open XN550 Drawer ", frame=F20_XN550_Draw, actionlist=[ActionManipulator.DRAWER_OPEN],
      | #         h_approach=p[0.07,0,0.1,0,0,0],
      | #         approach=p[0,0,0.1,0,0,0],
      | #         target = p[0,0,0,0,0,d2r(90)],
      | #         retract=p[0.07,0,0,0,0,0],
      | #         h_retract=p[0.07,0,0.1,0,0,0]
      | #         ))
      | # MOVEMENT_MAP.append(create_movement(description="Close XN550 Drawer ", frame=F20_XN550_Draw, actionlist=[ActionManipulator.DRAWER_CLOSE],
      | #         h_approach=p[0.07,0,0.1,0,0,0],
      | #         approach=p[0.07,0,0,0,0,0],
      | #         target = p[0,0,0,0,0,d2r(90)],
      | #         retract=p[0,0,0.1,0,0,0],
      | #         h_retract=p[0.07,0,0.1,0,0,0]
      | #         ))
      | # MOVEMENT_MAP.append(create_movement(description="Push XN550 Button ", frame=F21_XN550_Btn, actionlist=[ActionManipulator.PUSH],
      | #         approach=p[0,0,0.15,0,0,0],
      | #         retract=p[0,0,0.15,0,0,0]
      | #         ))
      | # MOVEMENT_MAP.append(create_movement(description="Capture Position 2 Input", frame=F_Cap_Input2,actionlist=[ActionManipulator.MOVE_TO]))
    Script file /programs/04 Scripts/SCRIPT Objects V0.1.script
      | #*****************************************************
      | # customer          :   INTERNAL
      | # project name      :
      | #****************************************************
      | # controller        :   UR
      | # software          :   5.17.3
      | #****************************************************
      | # author            :   P. Koehnke
      | # Copyright (c)     :   United Robotics Group
      | #                       An der Riede 2
      | #                       28816 Stuhr
      | #                       Germany
      | #****************************************************
      | # description       :   object database
      | # version:      	:   0.1
      | # created           :   09.10.2024
      | # updated           :
      | #****************************************************
      | # modifications     :
      | #
      | # date              :
      | # name              :
      | # reason            :
      | #****************************************************
      | 
      | def create_object_2(id=0, name="", type=0, dimension=struct(length=0, width=0, height=0, diameter=0), gripper_offset=p[0,0,0,0,0,0]):
      |     return struct(id=id, name=name, type=type, dimension=dimension, gripper_offset=gripper_offset)
      | end
      | 
      | OBJ = create_object_2()
      | OBJs = make_list(0, create_object_2(), 50)
      | 
      | OBJs.append(create_object_2(id=1, name="rack centrifuge", type=1, dimension=struct(length=0, width=0, height=0.106, diameter=0.020), gripper_offset=p[0,0,0.095,0,0,2.356]))
      | OBJs.append(create_object_2(id=2, name="sample tube 1", type=2, dimension=struct(length=0, width=0, height=0.106, diameter=0.015), gripper_offset=p[0,0,0,0,0,0]))
      | OBJs.append(create_object_2(id=3, name="rack sarstedt", type=3, dimension=struct(length=0, width=0, height=0.100, diameter=0.020), gripper_offset=p[0,0,0,0,0,0]))
      | OBJs.append(create_object_2(id=4, name="Lab bottle", type=4, dimension=struct(length=0, width=0, height=0.100, diameter=0.030), gripper_offset=p[0,0,0.2,0,0,0]))
      | OBJs.append(create_object_2(id=5, name="Vial", type=5, dimension=struct(length=0, width=0, height=0.100, diameter=0.0275), gripper_offset=p[0,0,0,0,0,0]))
      | OBJs.append(create_object_2(id=6, name="Container_S", type=6, dimension=struct(length=0.09, width=0.09, height=0.185, diameter=0.080), gripper_offset=p[0,0,0,0,0,0]))
      | OBJs.append(create_object_2(id=7, name="Target_container", type=7, dimension=struct(length=0.06, width=0.06, height=0.134, diameter=0.05), gripper_offset=p[0,0,0,0,0,0]))
      | OBJs.append(create_object_2(id=8, name="Spatula", type=8, dimension=struct(length=0.03, width=0.03, height=0.23, diameter=0.05), gripper_offset=p[0,0,0,0,0,0]))
      | OBJs.append(create_object_2(id=9, name="rack pipet", type=9, dimension=struct(length=0.03, width=0.03, height=0.23, diameter=0.05), gripper_offset=p[0,0,0,0,0,0]))
      | 
      | def create_jig_2(id=0, name="", type=0, capacity=0, jig_offset=p[0,0,0,0,0,0]):
      |     # iformation about used jigs
      |     return struct(id=id, name=name, type=type, capacity=capacity, jig_offset=jig_offset)
      | end
      | 
      | JIG2 = create_jig_2()
      | JIGs = make_list(0, create_jig_2(), 20)
      | 
      | JIGs.append(create_jig_2(id=1, name="3FG", type=1, capacity=1, jig_offset=p[0,0,0,0,0,0]))
      | JIGs.append(create_jig_2(id=2, name="jig input", type=2, capacity=1, jig_offset=p[0,0,0,0,0,-3.927]))
      | JIGs.append(create_jig_2(id=3, name="jig output", type=3, capacity=1, jig_offset=p[0,0,0,0,0,0.78]))
      | JIGs.append(create_jig_2(id=6, name="jig bin", type=6, capacity=1, jig_offset=p[0,0,0,0,0,0]))
      | JIGs.append(create_jig_2(id=7, name="jig sarstedt racks", type=7, capacity=1, jig_offset=p[0,0,-0.02,0,0,0]))
      | JIGs.append(create_jig_2(id=8, name="NoK Bin", type=8, capacity=1, jig_offset=p[0,0,0,0,0,0]))
      | JIGs.append(create_jig_2(id=9, name="Pick bott jig", type=9, capacity=1, jig_offset=p[0,0,0,0,0,0]))
      | JIGs.append(create_jig_2(id=10, name="Place bott jig", type=10, capacity=1, jig_offset=p[0,0,0,0,0,0]))
      | JIGs.append(create_jig_2(id=11, name="bottle shake jig", type=11, capacity=1, jig_offset=p[0,0,0,0,0,0]))
      | JIGs.append(create_jig_2(id=12, name="Pick Vial jig", type=12, capacity=1, jig_offset=p[0,0,0,0,0,0]))
      | JIGs.append(create_jig_2(id=13, name="Place Vial jig", type=13, capacity=1, jig_offset=p[0,0,0,0,0,0]))
      | JIGs.append(create_jig_2(id=14, name="Liquid transfer jig", type=14, capacity=1, jig_offset=p[0,0,0,0,0,0]))
      | JIGs.append(create_jig_2(id=15, name="Pick station jig", type=15, capacity=1, jig_offset=p[0,0,0,0,0,0]))
      | JIGs.append(create_jig_2(id=16, name="Place station jig", type=16, capacity=1, jig_offset=p[0,0,0,0,0,0]))
      | JIGs.append(create_jig_2(id=17, name="Weigh station jig", type=17, capacity=1, jig_offset=p[0,0,0,0,0,0]))
      | JIGs.append(create_jig_2(id=18, name="Pick station 1", type=18, capacity=1, jig_offset=p[0,0,0,0,0,0]))
      | JIGs.append(create_jig_2(id=19, name="Pick station 2", type=19, capacity=1, jig_offset=p[0,0,0,0,0,0]))
      | JIGs.append(create_jig_2(id=20, name="Pick station 3", type=20, capacity=1, jig_offset=p[0,0,0,0,0,0]))
      | JIGs.append(create_jig_2(id=21, name="Tilt station jig", type=21, capacity=1, jig_offset=p[0,0,0,0,0,0]))
    SuppressedNode
      Script file /programs/04 Scripts/krish.script
        | def vibration_2():
        | 	set_analog_out(0,0.4)
        | 	sleep(0.8)
        | 	set_analog_out(0,0.0)
        | 	sleep(0.2)
        | end
        | 
        | def vibration_3():
        | 	set_analog_out(0,0.4)
        | 	sleep(0.7)
        | 	set_analog_out(0,0.0)
        | 	sleep(0.3)
        | end
        | 
        | def vibration_4():
        | 	set_analog_out(0,0.4)
        | 	sleep(0.6)
        | 	set_analog_out(0, 0.0)
        | 	sleep(0.5)
        | end
        | 
        | def vibration_1():
        | 	set_analog_out(0,0.4)
        | 	sleep(1)
        | 	set_analog_out(0,0.0)
        | 	sleep(0)
        | end
        | 
        | def move_tilt_in_steps(PowA_center, final_pose, steps):
        | 	i = 0
        | 	while i <= steps:
        | 		ratio = i / steps
        | 		pose_step = p[PowA_center[0] + ratio * (final_pose[0] - PowA_center[0]), PowA_center[1] + ratio * (final_pose[1] -PowA_center[1]),PowA_center[2] + ratio * (final_pose[2] - PowA_center[2]), PowA_center[3] + ratio * (final_pose[3] - PowA_center[3]), PowA_center[4] + ratio * (final_pose[4] - PowA_center[4]), PowA_center[5] + ratio * (final_pose[5] - PowA_center[5])]
        | 		movej(pose_step, a=1.2, v=0.15)
        | 		sleep(0.1)
        | 		i = i+1
        | 	end
        | end
        | 
        | def tilt_container(angle):
        | 	P_center = get_actual_tcp_pose()
        | 	hinge_offset = p[0,0,-0.23,0,0,0]
        | 	pivot_pose = pose_trans(P_center, hinge_offset)
        | 	pose_rel = pose_trans(pose_inv(pivot_pose), P_center)
        | 	angle_mid = (angle/2.0)*3.1416/180
        | 	angle_end = angle*3.1416/180
        | 	tilt_mid = p[0,0,0, -angle_mid, 0, 0]
        | 	tilt_end = p[0,0,0, -angle_end, 0, 0]
        | 	pose_rel_mid = pose_trans(tilt_mid, pose_rel)
        | 	pose_rel_end = pose_trans(tilt_end, pose_rel)
        | 	via_pose = pose_trans(pivot_pose, pose_rel_mid)
        | 	end_pose = pose_trans(pivot_pose, pose_rel_end)
        | 	movec(via_pose, end_pose, a=0.05, v=0.01, r=0.001)
        | 	P_center = get_actual_tcp_pose()
        | end
        | 
        | def deg2rad(d):
        | 	return d*3.141592/180
        | end
        | 
        | def map_tilt_to_ry_deg(container_deg):
        | 	#ry_deg = -0.875*container_deg +87.0
        | 	#return clamp(ry_deg, 5.0, 80.0)
        | 	if (Pow_name == "NaCl" or Pow_name == "Mannitol" or Pow_name == "CCS" or Pow_name == "lactose_loose"):
        | 		if ( level>=10.0):
        | 			ry_min = 10.0
        | 			ry_max = 75.0
        | 		elif (level<10.00 and level >1.00):
        | 			ry_min = 16.0
        | 			ry_max = 65.0
        | 		else:
        | 			ry_min=17.0
        | 			ry_max=75.0
        | 		end
        | 	else:
        | 		if ( level>=10.0):
        | 			ry_min = 0.0
        | 			ry_max = 55.0
        | 		elif (level<10.00 and level >1.00):
        | 			ry_min = 10.0
        | 			ry_max = 45.0
        | 		else:
        | 			ry_min=0.0
        | 			ry_max=50.0
        | 		end
        | 
        | 	end
        | 	local span_count = angle_max -angle_min
        | 	local span_ry = ry_max - ry_min
        | 
        | 	local t = (container_deg -angle_min)/span_count
        | 	local ry_deg = ry_max - t*span_ry
        | 
        | 	return clamp(ry_deg, ry_min, ry_max)
        | 
        | end
        | 
        | def caluclate_corrections(level):
        | 	z_high = 0.01
        | 	z_low = -0.08
        | 	y_high = -0.010
        | 	y_low = -0.03
        | 
        | 	scale = (level - 10.0) / (100.0-10.0)
        | 
        | 	global correction_z = z_low + scale*(z_high - z_low)
        | 	global correction_y = y_low + scale*(y_high -y_low)
        | 
        | end
        | 
        | def scoop_powder(P_center):
        | 	#lift_offset = p[0, 0, 0.05, 0, 0, 0]
        | 	vibration_voltage = 0.4
        | 	vibration_time = 3.0
        | 	diameter = 0.07
        | 	global scoop_radius_default = 0.0
        | 	#P_center = center_pose_t
        | 
        | 
        | 	if (level >=70.00):
        | 		approach_offset = p[0.008,0,0.22,0,0,0]
        | 		lift_offset = p[0, 0, 0.12, 0, 0, 0]
        | 		caluclate_corrections(level)
        | 	elif (level >=10.00 and level <70):
        | 		approach_offset = p[0.008,0,0.22,0,0,0]
        | 		lift_offset = p[0, 0, 0.15, 0, 0, 0]
        | 		caluclate_corrections(level)
        | 	elif (level<10.00 and level >= 1.00):
        | 		approach_offset = p[0.006,0,0.22,0,0,0]
        | 		correction_z = -0.08
        | 		correction_y = -0.01
        | 		lift_offset = p[0, 0, 0.14, 0, 0, 0]
        | 	else:
        | 		approach_offset = p[0.008,0,0.22,0,0,0]
        | 		correction_z = -0.08
        | 		correction_y = -0.01
        | 		lift_offset = p[0, 0, 0.14, 0, 0, 0]
        |  	end
        | 
        | 	if (spatula == "spatula_L"):
        | 		global spatula_depth = 0.015
        | 	elif (spatula == "spatula_M"):
        | 		global spatula_depth = 0.01
        | 	elif (spatula == "spatula_S"):
        | 		global spatula_depth = 0.006
        | 	elif (spatula == "spatula_flat_M"):
        | 		global spatula_depth = 0.001
        | 	elif (spatula == "spatula_flat_S"):
        | 		global spatula_depth = 0.005
        | 	end
        | 
        | 	scoop_radius_default = diameter/2 - spatula_depth
        | 	scoop_entry_pose = pose_trans(P_center, approach_offset)
        | 	movel(scoop_entry_pose, a=0.05, v=0.05)
        | 
        | 	scoop_start_rel = p[scoop_radius_default, 0, scoop_depth, 0, 0, 0]
        | 
        | 	rot_mid = p[0, 0, 0, 0, 0, 0.785]
        | 	rot_end = p[0, 0, 0, 0, 0, 1.5708]
        | 
        | 	scoop_via_rel = pose_trans(rot_mid, scoop_start_rel)
        | 	scoop_end_rel = pose_trans(rot_end, scoop_start_rel)
        | 
        | 	scoop_start_pose = pose_trans(P_center, scoop_start_rel)
        | 	scoop_via_pose = pose_trans(P_center, scoop_via_rel)
        | 	scoop_end_pose = pose_trans(P_center, scoop_end_rel)
        | 
        | 	movel(scoop_start_pose, a=0.3, v=0.7)
        | 
        | 	if (level<90.0):
        | 		Rotate()
        | 	end
        | 
        | 	#movec(scoop_via_pose, scoop_end_pose, a=0.03, v=0.05)
        | 	movec(scoop_via_pose, scoop_end_pose, a=0.03, v=0.02)
        | 	#movel(pose_trans(get_actual_tcp_pose(), p[0,0,0,0,0,deg2rad(90.0)]), a=0.03, v=0.05)
        | 	sleep(1.0)
        | 	local ry_deg = map_tilt_to_ry_deg(angle_deg)
        | 	local ry = deg2rad(ry_deg)
        | 	local end_rel = pose_trans(pose_inv(P_center), scoop_end_pose)
        | 	local end_rel_tilted = pose_trans(end_rel, p[0, 0, 0, 0, ry, 0])
        | 	global tilted_pose_in_base = pose_trans(P_center, p[0,correction_y,correction_z,end_rel_tilted[3],end_rel_tilted[4], end_rel_tilted[5]])
        | 	global tilted_pose_in_base = pose_trans(tilted_pose_in_base, p[0, 0, spatula_len, 0, 0, 0])
        | 
        | 	movel(tilted_pose_in_base, a=0.03, v=0.1)
        | 	set_analog_out(0, vibration_voltage)
        | 
        | 	local ry_level = deg2rad(ry_deg/1.5)
        | 	local end_rel_tilted_level = pose_trans(end_rel, p[0, 0, 0, 0, ry_level, 0])
        | 	local level_tilted_pose_in_base = pose_trans(P_center, p[0,correction_y,correction_z,end_rel_tilted_level[3],end_rel_tilted_level[4], end_rel_tilted_level[5]])
        | 	local level_tilted_pose_in_base = pose_trans(level_tilted_pose_in_base, p[0, 0, spatula_len, 0, 0, 0])
        | 
        | 	movel(level_tilted_pose_in_base, a=0.03, v=0.1)
        | 	#if (level>70.0):
        | 		#sleep(1.0)
        | 	#end
        | 	sleep(2.0)
        | 	#sleep(vibration_time)
        | 
        | 	movel(tilted_pose_in_base, a=0.03, v=0.1)
        | 	set_analog_out(0, 0.0)
        | 
        | 	tilt_pose_rel = pose_trans(pose_inv(P_center), tilted_pose_in_base)
        | 
        | 	lifted_pose_rel = pose_trans(lift_offset, tilt_pose_rel)
        | 
        | 	global lifted_pose = pose_trans(P_center, lifted_pose_rel)
        | 	movel(lifted_pose, a=0.03, v=0.1)
        | end
        | 
        | 
        | def center_pose():
        | 	trans_rel = p[-0.014, 0.06, -0.015, 0, 0, 0]
        | 
        | 	p_translated = pose_trans(place_pose, trans_rel)
        | 	cx = p_translated[0]
        | 	cy = p_translated[1]
        | 	cz = p_translated[2]
        | 
        | 	global P_center_vertical = p[cx,cy,cz, 0, 0, 4.08]
        | 
        | 	#movej(P_center_vertical, a =0.3, v =0.3)
        | 	return P_center_vertical
        | end
        | 
        | def updated_center_pose(P_center_vertical, angle_deg):
        | 	hinge_pose = pose_trans(P_center_vertical, p[0,0,-0.2,0,0,0])
        | 	local_rel = pose_trans(pose_inv(hinge_pose), P_center_vertical)
        | 
        | 	rot_tilt = p[0,0,0, -deg2rad(angle_deg),0,0]
        | 	local_rel_tilted = pose_trans(rot_tilt, local_rel)
        | 
        | 	global P_center = pose_trans(hinge_pose, local_rel_tilted)
        | 	return P_center
        | end
        | 
        | def tilt_send(angle):
        | 	socket_open("192.168.12.105", 80)
        | 	angle = 85.0 - angle
        | 	socket_send_string("Tilt,"+to_str(angle)+",0")
        | 	sync()
        | 	sleep(0.5)
        | 	socket_close()
        | end
        | 
        | def Motors_off():
        | 	socket_open("192.168.12.105", 80)
        | 	socket_send_string("Off,0,0")
        | 	sync()
        | 	sleep(0.5)
        | 	socket_close()
        | end
        | 
        | def Rotate():
        | 	socket_open("192.168.12.105", 80)
        | 	socket_send_string("FullRotation, 1, 2000")
        | 	sync()
        | 	sleep(0.5)
        | 	socket_close()
        | end
        | 
        | def tilt_to_home():
        | 	socket_open("192.168.12.105", 80)
        | 	socket_send_string("Home,0,0")
        | 	sync()
        | 	sleep(0.5)
        | 	socket_close()
        | end
  Folder BeforeStarts [hidden by the author, left out]
Robot Program (runOnlyOnce=false)
  Folder MAIN
    Script: command_manager(external_control="uGO", cond_suspend=(ITM_Manipulated and AMR_AtTarget and AMR_Charging and AMR_Battery<40), cond_unsuspend=(AMR_Battery≟60))
    Script: log_state(STATE_Info)
    Switch expression=STATE
      Case (caseValue=1)
        Folder Stopping
          STATE_Info := "Stopping"
          Script: end_freedrive_mode()
          Set NoAction tcp=TCP
          PSE_T := get_tool_free_pose(dir=[0,0,0.150], move_in_base_frame=True)
          If is_reachable(Base, [PSE_T])
            MoveL speed 150 mm/s, acceleration 1200 mm/s^2 (useActiveTCP=true) feature=Base
              Waypoint Variable (Variable): variable=PSE_T
          Script: do_transition(keep_rxry=OBJ_Picked, r=0)
          SuppressedNode
            Folder Decapper
              Set DigitalOutput pin=digital_out[4]; digitalValue=0
              Set DigitalOutput pin=BarcodeTrigger; digitalValue=0
              Set DigitalOutput pin=digital_out[3]; digitalValue=0
              Set DigitalOutput pin=digital_out[2]; digitalValue=0
              Set DigitalOutput pin=digital_out[5]; digitalValue=0
          SuppressedNode
            Folder Centrifuge [hidden by the author, left out]
          Call Sub_AMR_MiR_V3
          If stopping() and AMR_Done
            STATE := 2
            Script: ugo_update_outputs()
      Case (caseValue=2)
        Folder Stopped [hidden by the author, left out]
      Case (caseValue=3)
        Folder  Resetting [hidden by the author, left out]
      Case (caseValue=4)
        Folder Idle [hidden by the author, left out]
      Case (caseValue=5)
        Folder Starting
          STATE_Info := "Starting"
          'ADD COMMANDS WHAT TO START WITH'
          Call Sub_AMR_MiR_V3
          Folder get ugo data
            Folder Assign Tasks
              Script: TASK.ID = ugo_get_task()
              If TASK.ID≟1
                Task_info := "Charge"
                Folder Parameters
                  AMR_PosTarget := 1
              ElseIf TASK.ID≟9
                'Pick Sarstedt Rack from Variable source'
                Task_info := "Navigate to Target"
                Folder Parameters
                  AMR_PosTarget := UGO.read_input("00","ITM_ID")
              ElseIf TASK.ID≟10
                'Pick Sarstedt Rack from Variable source'
                Task_info := "Pick Rack"
                AMR_PosTarget := 2
                Folder Parameters
                  ITM_ID := UGO.read_input("00","ITM_ID")
                  JIG := UGO.read_input("00","JIG_ID")
                  OBJ_Type := 3
              ElseIf TASK.ID≟11
                'Place Sarstedt Rack on Variable target'
                Task_info := "Place Rack"
                AMR_PosTarget := 2
                Folder Parameters [hidden by the author, left out]
                SuppressedNode
                  ITM_ID := 1
              ElseIf TASK.ID≟12
                Task_info := "Decapping"
                Folder Parameters
                  ITM_ID := 1
                  AMR_PosTarget := AMR_PosActual
                  PRC_TubCounter := 0
              ElseIf TASK.ID≟13
                Task_info := "Empty racks"
                Folder Parameters [hidden by the author, left out]
              ElseIf TASK.ID≟16
                Task_info := "Decap + Barcode"
                Folder Parameters [hidden by the author, left out]
              ElseIf TASK.ID≟30
                Task_info := "Getting bottles"
                Folder Parameters
                  ITM_ID := 1
                  OBJ_Type := 4
                  JIG := 9
                  AMR_PosTarget := 4
              ElseIf TASK.ID≟40
                Task_info := "Placing bottles"
                Folder Parameters
                  ITM_ID := 1
                  OBJ_Type := 4
                  JIG := 10
                  AMR_PosTarget := 4
              ElseIf TASK.ID≟41
                Task_info := "Shaking bottle"
                Folder Parameters
                  ITM_ID := 1
                  OBJ_Type := 4
                  JIG := 11
                  AMR_PosTarget := 4
              ElseIf TASK.ID≟42
                Task_info := "Decap the bottle"
                Folder Parameters
                  ITM_ID := 1
                  OBJ_Type := 4
                  AMR_PosTarget := 4
              ElseIf TASK.ID≟43
                Task_info := "Pick the Rack"
                AMR_PosTarget := 5
                Folder Parameters
                  ITM_ID := UGO.read_input("00","ITM_ID")
                  JIG := UGO.read_input("00","JIG_ID")
                  OBJ_Type := 3
              ElseIf TASK.ID≟45
                Task_info := "pick the Vial"
                Folder Parameters
                  ITM_ID := 1
                  OBJ_Type := 4
                  JIG := 12
                  AMR_PosTarget := 5
              ElseIf TASK.ID≟46
                Task_info := "Decap the Vial"
                Folder Parameters
                  ITM_ID := 1
                  OBJ_Type := 4
                  JIG := 13
                  AMR_PosTarget := 5
              ElseIf TASK.ID≟47
                Task_info := "Liquid Transfer"
                Folder Parameters
                  ITM_ID := 1
                  OBJ_Type := 4
                  JIG := 14
                  AMR_PosTarget := 3
              ElseIf TASK.ID≟48
                Task_info := "Place_rack"
                Folder Parameters
                  ITM_ID := 1
                  OBJ_Type := 3
                  JIG := 7
                  AMR_PosTarget := 5
              ElseIf TASK.ID≟49
                Task_info := "Pick Containers"
                Folder Parameters
                  ITM_ID := 1
                  OBJ_Type := 6
                  JIG := 15
                  AMR_PosTarget := 3
              ElseIf TASK.ID≟50
                Task_info := "Decap Containers"
                Folder Parameters
                  ITM_ID := 1
                  OBJ_Type := 6
                  JIG := 16
                  AMR_PosTarget := 5
              ElseIf TASK.ID≟51
                Task_info := "Detect Spatula and transfer powder"
                Folder Parameters
                  ITM_ID := 1
                  OBJ_Type := 8
                  JIG := 16
                  AMR_PosTarget := 5
              ElseIf TASK.ID≟99
                Task_info := "Decapping and barcode alignment"
                Folder Parameters
                  PRC_TubNumber := UGO.read_input("00","TubesNb")
                  PRC_TubCounter := 0
                  ITM_ID := 1
                  AMR_PosTarget := AMR_PosActual
              SuppressedNode
                ElseIf TASK.ID≟14
                  Task_info := "Load Centrifuge"
                  Folder Parameters
                    PRC_RackCounter := 0
                    Script: TASK.WORK.ITM_ID_Src=1
                    Script: TASK.WORK.ITM_ID_Tgt=2
                    AMR_PosTarget := 4
                    AMR_FootprintID := 1
              SuppressedNode
                ElseIf TASK.ID≟15
                  Task_info := "Unoad Centrifuge"
                  Folder Parameters [hidden by the author, left out]
              SuppressedNode
                ElseIf TASK.ID≟99
                  Task_info := "Load Biorad"
                  Folder Parameters
                    PRC_RackCounter := 0
                    ITM_ID := 2
                    CAM_LM_ID := 0
                    SuppressedNode
                      AMR_PosTarget := 1
                    AMR_PosTarget := AMR_PosActual
                    PRC_RackNumber := UGO.read_input("00","RackNb")
              SuppressedNode
                ElseIf TASK.ID≟99
                  Task_info := "Unload Biorad"
                  Folder Parameters
                    PRC_RackCounter := 0
                    ITM_ID := 2
                    CAM_LM_ID := 0
                    SuppressedNode
                      AMR_PosTarget := 1
                    AMR_PosTarget := AMR_PosActual
                    PRC_RackNumber := UGO.read_input("00","RackNb")
              Else 
                Script: set_error(ERROR_WRONG_ORDER)
          Folder test ugo
            Wait Sleep waitTime=0.2
            Script: ugo_update_outputs()
          If starting() and AMR_Done
            Script: log_message(Task_info, "New Task: ")
            Script: log_message(to_str(TASK.ID), "Task_ID: ")
            Script: do_transition(keep_rxry=OBJ_Picked)
            STATE := 6
            Script: ugo_update_outputs()
      Case (caseValue=6)
        Folder Execute
          STATE_Info := "Execute"
          If not CMD_Hold and not CMD_Suspend (checkContinuously=true)
            Switch expression=PROCESS_Step
              Case (caseValue=0)
                PROCESS_Info := "process control"
                Script: log_process(PROCESS_Info)
                Folder process control [hidden by the author, left out]
              Case (caseValue=1)
                Folder navigate [hidden by the author, left out]
              Case (caseValue=2)
                Folder prepare [hidden by the author, left out]
              Case (caseValue=3)
                Folder work
                  'ADD EVERY MACHINE, OBJECT, STATION TO WORK ON'
                  Switch expression=ITM_ID
                    Case (caseValue=1)
                      Folder uLM
                        If TASK.ID≟12
                          Folder fill racks
                            Action := 151
                            Call Sub_Vision_V18
                            If not ERROR.FLAG
                              Folder Actions for the task
                                Action := 1
                                JIG := 2
                                JIG_Slot := CAM_Result[0]
                                OBJ_Nbr := CAM_Result[0]
                                OBJ_Type := 2
                                Call Sub_Action_V4
                                If OBJ_Picked
                                  Script: CAM_Result.remove(0)
                                  PRC_TubCounter := PRC_TubCounter+1
                                  If PRC_TubCounter%4≟0
                                    JIG_Slot := 4
                                  Else 
                                    JIG_Slot := PRC_TubCounter%4
                                  OBJ_Nbr := ceil(PRC_TubCounter/4)
                                  Action := 2
                                  JIG := 4
                                  Call Sub_Action_V4
                                  Action := 151
                                  Call Sub_Vision_V18
                            If (CAM_Captures≥CAM_PRM_Retries) or (PRC_TubCounter≥32)
                              PROCESS_Step := 0
                              WRK_Done := True
                        ElseIf TASK.ID≟10
                          Folder Pick Rack
                            Action := 131
                            Call Sub_Vision_V18
                            Action := 1
                            Call Sub_Action_V4
                            PROCESS_Step := 0
                            WRK_Done := True
                        ElseIf TASK.ID≟11
                          Folder Place Rack [hidden by the author, left out]
                        ElseIf TASK.ID≟13
                          Folder empty racks
                            Folder pick
                              Action := 1
                              JIG := 4
                              If PRC_TubCounter%4≟0
                                JIG_Slot := 4
                              Else 
                                JIG_Slot := PRC_TubCounter%4
                              OBJ_Nbr := ceil(PRC_TubCounter/4)
                              OBJ_Type := 2
                              Call Sub_Action_V4
                              If OBJ_Picked
                                Action := 2
                                JIG := 3
                                JIG_Slot := 1
                                CNT_Rack_Output := CNT_Rack_Output + 1
                                OBJ_Nbr := CNT_Rack_Output
                                Call Sub_Action_V4
                                If not ERROR.FLAG
                                  PRC_TubCounter := PRC_TubCounter - 1
                              If CNT_Rack_Output≥50 or PRC_TubCounter≤0
                                PROCESS_Step := 0
                                WRK_Done := True
                        ElseIf TASK.ID≟16
                          CAM_Result := OBJs_List
                          PRC_CntDetect := 0
                          Loop While (checkContinuously=false) expression=PRC_CntDetect<CAM_Result.length()
                            Action := 1
                            ITM_ID := 1
                            JIG := 2
                            OBJ_Type := 2
                            JIG_Slot := CAM_Result[PRC_CntDetect]
                            OBJ_Nbr := CAM_Result[PRC_CntDetect]
                            Call Sub_Action_V4
                            JIG := 1
                            Action := 11
                            Call Sub_Action_V4
                            Action := 12
                            Call Sub_Action_V4
                            Action := 6
                            JIG := 6
                            Call Sub_Action_V4
                            Action := 13
                            Call Sub_Action_V4
                            Action := 1
                            JIG := 1
                            Call Sub_Action_V4
                            If OBJ_Brc_OK
                              JIG := 2
                              Action := 2
                              OBJ_Nbr := CAM_Result[PRC_CntDetect]
                              JIG_Slot := CAM_Result[PRC_CntDetect]
                              OBJ_Type := 2
                              Call Sub_Action_V4
                            Else 
                              Action := 2
                              JIG := 8
                              Call Sub_Action_V4
                            PRC_CntDetect := PRC_CntDetect+1
                          PROCESS_Step := 0
                          WRK_Done := True
                        ElseIf TASK.ID≟30
                          Folder Pick Bottle
                            Action := 1
                            Call Sub_Action_V4
                            PROCESS_Step := 0
                            WRK_Done := True
                        ElseIf TASK.ID≟40
                          Folder Place Bottle
                            Action := 2
                            Call Sub_Action_V4
                            PROCESS_Step := 0
                            WRK_Done := True
                        ElseIf TASK.ID≟45
                          Folder Pick Vial
                            Action := 31
                            Call Sub_Action_V4
                            PROCESS_Step := 0
                            WRK_Done := True
                        ElseIf TASK.ID≟46
                          Folder Decap Vial
                            Action := 32
                            Call Sub_Action_V4
                            PROCESS_Step := 0
                            WRK_Done := True
                        ElseIf TASK.ID≟47
                          Folder Liquid transfer
                            Action := 33
                            Call Sub_Action_V4
                            PROCESS_Step := 0
                            WRK_Done := True
                        ElseIf TASK.ID≟48
                          Folder Place Rack
                            Action := 34
                            Call Sub_Action_V4
                            PROCESS_Step := 0
                            WRK_Done := True
                        ElseIf TASK.ID≟49
                          Folder Pick Powder container
                            Action := 35
                            Call Sub_Action_V4
                            PROCESS_Step := 0
                            WRK_Done := True
                        ElseIf TASK.ID≟41
                          Folder shake Bottle
                            Action := 30
                            Call Sub_Action_V4
                            PROCESS_Step := 0
                            WRK_Done := True
                        ElseIf TASK.ID≟42
                          Folder decap the bottle
                            Action := 1
                            JIG := 9
                            Call Sub_Action_V4
                            Action := 11
                            JIG := 1
                            Call Sub_Action_V4
                            Action := 12
                            JIG := 1
                            Call Sub_Action_V4
                            Action := 2
                            JIG := 8
                            Call Sub_Action_V4
                            PROCESS_Step := 0
                            WRK_Done := True
                        ElseIf TASK.ID≟43
                          Folder Pick the rack
                            Action := 131
                            Call Sub_Vision_V18
                            Action := 1
                            Call Sub_Action_V4
                            PROCESS_Step := 0
                            WRK_Done := True
                        ElseIf TASK.ID≟50
                          Folder Decap containers
                            Action := 36
                            Call Sub_Action_V4
                            PROCESS_Step := 0
                            WRK_Done := True
                        ElseIf TASK.ID≟51
                          Folder Detect Spatula and transfer powder
                            Action := 37
                            Call Sub_Action_V4
                            PROCESS_Step := 0
                            WRK_Done := True
                    Case (caseValue=2)
                      SuppressedNode
                        Folder Centrfiuge
                          SuppressedNode
                            Script: cent_error_check()
                          OBJ_Type := 1
                          If not ERROR.FLAG
                            'load racks'
                            If TASK.ID≟14
                              Loop While (checkContinuously=false) expression=(PRC_RackCounter<4) and  not CMD_Stop and  not ERROR.FLAG
                                ITM_ID := TASK.WORK.ITM_ID_Src
                                JIG := 4
                                JIG_Slot := PRC_RackCounter+1
                                Action := 1
                                Call Sub_Action_V4
                                If OBJ_Picked and  not ERROR.FLAG
                                  ITM_ID := TASK.WORK.ITM_ID_Tgt
                                  Script: execute_cent_action(ACTION_ROTATE, JIG_Slot)
                                  Action := 7
                                  Call Sub_Action_V4
                                  PRC_RackCounter := PRC_RackCounter + 1
                              If not ERROR.FLAG
                                WRK_Done := True
                                PROCESS_Step := 0
                            'unload racks'
                            If TASK.ID≟15
                              If CNT_State_Actual≟2 or CNT_State_Actual≟3
                                Loop While (checkContinuously=false) expression=(PRC_RackCounter<4) and  not CMD_Stop and  not ERROR.FLAG
                                  ITM_ID := TASK.WORK.ITM_ID_Src
                                  JIG_Slot := PRC_RackCounter + 1
                                  Script: execute_cent_action(ACTION_ROTATE, JIG_Slot)
                                  Script: execute_cent_action(ACTION_INSPECT, JIG_Slot)
                                  Action := 8
                                  Call Sub_Action_V4
                                  If OBJ_Picked and  not ERROR.FLAG
                                    ITM_ID := TASK.WORK.ITM_ID_Tgt
                                    JIG := 4
                                    JIG_Slot := PRC_RackCounter + 1
                                    Action := 2
                                    Call Sub_Action_V4
                                    PRC_RackCounter := PRC_RackCounter+1
                                If not ERROR.FLAG
                                  WRK_Done := True
                                  PROCESS_Step := 0
                    Case (caseValue=5)
                      Folder SarstedtTable
                        Action := 131
                        Call Sub_Vision_V18
                        Action := 1
                        Call Sub_Action_V4
                        PROCESS_Step := 0
                        WRK_Done := True
                    Case (caseValue=20)
                      SuppressedNode
                        Folder Biorad rack
                          'load racks'
                          If Task_ID≟16
                            SuppressedNode
                              PRC_RackCounter := 0
                            Loop While (checkContinuously=false) expression=(PRC_RackCounter<PRC_RackNumber) and  not CMD_Stop
                              JIG_Slot := PRC_RackCounter
                              Action := 1
                              PRC_Target := 0
                              Call Sub_Action_V4
                              If OBJ_Picked
                                Action := 2
                                PRC_Target := 1
                                Call Sub_Action_V4
                                Action := 7
                                PRC_Target := 1
                                Call Sub_Action_V4
                                PRC_RackCounter := PRC_RackCounter+1
                            WRK_Done := True
                            PROCESS_Step := 0
                          'unload racks'
                          SuppressedNode
                            If Task_ID≟17
                              SuppressedNode
                                PRC_RackCounter := 0
                              Loop While (checkContinuously=false) expression=(PRC_RackCounter<PRC_RackNumber) and  not CMD_Stop
                                JIG_Slot := PRC_RackCounter
                                Action := 8
                                PRC_Target := 1
                                Script: textmsg("Callactionunload=",Action)
                                Call Sub_Action_V4
                                Action := 1
                                PRC_Target := 1
                                Script: textmsg("Callactionpick=",Action)
                                Call Sub_Action_V4
                                If OBJ_Picked
                                  Action := 2
                                  PRC_Target := 0
                                  Script: textmsg("Callactionplace=",Action)
                                  Call Sub_Action_V4
                                  PRC_RackCounter := PRC_RackCounter+1
                              WRK_Done := True
                              PROCESS_Step := 0
                          If Task_ID≟17
                            PRC_RackCounter := 0
                            Loop While (checkContinuously=false) expression=(PRC_RackCounter<PRC_RackNumber) and  not CMD_Stop
                              Wait Condition expression=SensorData[PRC_RackCounter]≟1
                              JIG_Slot := PRC_RackCounter
                              Action := 8
                              PRC_Target := 1
                              Script: textmsg("Callactionunload=",Action)
                              Call Sub_Action_V4
                              Action := 1
                              PRC_Target := 1
                              Script: textmsg("Callactionpick=",Action)
                              Call Sub_Action_V4
                              If OBJ_Picked
                                Action := 2
                                PRC_Target := 0
                                Script: textmsg("Callactionplace=",Action)
                                Call Sub_Action_V4
                                PRC_RackCounter := PRC_RackCounter+1
                            WRK_Done := True
                            PROCESS_Step := 0
                    Case (caseValue=43)
                      Folder Pick the rack
                        Action := 131
                        Call Sub_Vision_V18
                        Action := 1
                        Call Sub_Action_V4
                        PROCESS_Step := 0
                        WRK_Done := True
                    Case (caseValue=2147483647)
                      WRK_Done := True
                      PROCESS_Step := 0
          If CMD_Hold
            STATE := 9
            Script: ugo_update_outputs()
          ElseIf CMD_Suspend
            STATE := 12
            Script: ugo_update_outputs()
      Case (caseValue=7)
        Folder Completing [hidden by the author, left out]
      Case (caseValue=8)
        Folder Complete [hidden by the author, left out]
      Case (caseValue=9)
        Folder Holding [hidden by the author, left out]
      Case (caseValue=10)
        Folder Held [hidden by the author, left out]
      Case (caseValue=11)
        Folder Unholding [hidden by the author, left out]
      Case (caseValue=12)
        Folder Suspending [hidden by the author, left out]
      Case (caseValue=13)
        Folder Suspended [hidden by the author, left out]
      Case (caseValue=14)
        Folder Unsuspending [hidden by the author, left out]
      Case (caseValue=15)
        Folder Aborting [hidden by the author, left out]
      Case (caseValue=16)
        Folder Aborted [hidden by the author, left out]
      Case (caseValue=17)
        Folder Clearing [hidden by the author, left out]
    Script: log_state(STATE_Info)
    Script: log_warning(WARNING.MSG)
    Script: log_error(ERROR.MSG)
    Folder Times [hidden by the author, left out]
    SuppressedNode
      Script: sync()
    Wait Sleep waitTime=0.1
SuppressedNode
  Thread Thread_1 (runOnlyOnce=false)
    Wait Condition expression=decap≟ True
    Set DigitalOutput pin=GRP_3F_Enable; digitalValue=1
    Set DigitalOutput pin=GRP_3F_Decap; digitalValue=1
    Wait Condition expression=decap≟ False
    Set DigitalOutput pin=GRP_3F_Enable; digitalValue=0
    Set DigitalOutput pin=GRP_3F_Decap; digitalValue=0
    Script: sync()
SubProgram -> Sub_Vision_V18
SubProgram  [hidden by the author, left out]
SubProgram -> Sub_Action_V4
SubProgram Sub_AMR_MiR_V3 [hidden by the author, left out]
SubProgram Sub_Action_V4 (keepSynchronizedWithDisk=true) programFile=/programs/03 Sub Routines/Sub_Action_V4.urp
  Folder PreSettings
    Folder init poses [hidden by the author, left out]
    Folder Gripping parameters [hidden by the author, left out]
    Switch expression=ITM_ID
      Case (caseValue=1)
        Folder uML
          Script: JIG2 = find_object_by_type(JIGs, JIG)
          JIG_Offset := JIG2.jig_offset
          Switch expression=JIG
            Case (caseValue=1)
              Folder 3FG
                Folder define poses
                  FRM_Reference := ULM_3FG
                  JNT_Q := JNT_HOME
                  PSE_T := pose_trans(GRP_Offset, JIG_Offset)
                  PSE_A := pose_trans(PSE_T, p[0,0,0.100,0,0,0])
                  PSE_R := pose_add(PSE_T, p[0,0,0.100,0,0,0])
            Case (caseValue=2)
              Folder Input
                'CHANGE THE REFERENCE TO THE FRAME TO MOVE IN'
                Folder define poses
                  FRM_Reference := ULM_Input
                  PSE_T := pose_trans(pose_trans(get_pattern_pos_rectangle(OBJ_Nbr, "X", [10,5], patternsize=[0.181,0.081]), GRP_Offset), JIG_Offset)
                  If Action≟1
                    PSE_R := pose_add(PSE_T, p[0,0,0.200,0,0,0])
                    PSE_A := pose_add(PSE_T, p[0,0,0.100,0,0,0])
                  ElseIf Action≟2
                    PSE_R := pose_add(PSE_T, p[0,0,0.100,0,0,0])
                    PSE_A := pose_add(PSE_T, p[0,0,0.200,0,0,0])
            Case (caseValue=3)
              Folder Output [hidden by the author, left out]
            Case (caseValue=4)
              Folder jig centrifuge racks [hidden by the author, left out]
            Case (caseValue=6)
              Folder Caps bin
                Folder define poses
                  'Drop cap'
                  Script: FRM_Reference=ULM_Cap_Bin
                  PSE_T := pose_RPY2RotVec(p[0,0,0,0,0,0])
                  PSE_T_H := pose_add(PSE_T, p[0,0,-0.011,0,0,0])
                  PSE_A := pose_trans(PSE_T, p[0,0,0.1,0,0,0])
                  PSE_R_H := pose_add(PSE_T, p[0,0,0.100,0,0,0])
                  PSE_R := pose_add(PSE_T, p[0,0,0.100,0,0,0])
            Case (caseValue=7)
              Folder Sarstedt [hidden by the author, left out]
            Case (caseValue=8)
              Folder NoK
                Folder define poses
                  'NoK'
                  Script: FRM_Reference=ULM_NoK
                  PSE_T := pose_RPY2RotVec(p[0,0,0,0,0,0])
                  PSE_A := pose_trans(PSE_T, p[0,0,0.1,0,0,0])
                  PSE_R := pose_add(PSE_T, p[0,0,0.100,0,0,0])
            Case (caseValue=9)
              Folder Pick_bott_jig
                Folder define poses
                  'NoK'
                  Script: FRM_Reference=ULM_bottle_pick
                  PSE_T := pose_RPY2RotVec(p[0,0,0,0,0,0])
                  PSE_A := pose_trans(PSE_T, p[0,0,0.1,0,0,0])
                  PSE_R := pose_add(PSE_T, p[0,0,0.100,0,0,0])
            Case (caseValue=10)
              Folder Place_bott_jig
                Folder define poses
                  'NoK'
                  Script: FRM_Reference=ULM_bottle_plac
                  PSE_T := pose_RPY2RotVec(p[0,0,0,0,0,0])
                  PSE_A := pose_trans(PSE_T, p[0,0,0.1,0,0,0])
                  PSE_R := pose_add(PSE_T, p[0,0,0.100,0,0,0])
            Case (caseValue=11)
              Folder Place_bott_jig
                Folder define poses
                  'NoK'
                  Script: FRM_Reference=shake
                  PSE_T := pose_RPY2RotVec(p[0,0,0,0,0,0])
                  PSE_A := pose_trans(PSE_T, p[0,0,0,0,0,0])
                  PSE_R := pose_add(PSE_T, p[0,0,0,0,0,0])
            Case (caseValue=12)
              Folder Pick_Vial_jig
                Folder define poses
                  'NoK'
                  Script: FRM_Reference=shake
                  PSE_T := pose_RPY2RotVec(p[0,0,0,0,0,0])
                  PSE_A := pose_trans(PSE_T, p[0,0,0,0,0,0])
                  PSE_R := pose_add(PSE_T, p[0,0,0,0,0,0])
      Case (caseValue=2)
        Folder Centrifuge
          'CHANGE THE REFERENCE TO THE FRAME TO MOVE IN'
          Folder define poses
            FRM_Reference := FRM_Centrifuge
            PSE_T := GRP_Offset
            If Action≟8
              PSE_R := pose_add(PSE_T, p[0,0,0.250,0,0,0])
              PSE_A := pose_add(PSE_T, p[0,0,0.150,0,0,0])
            ElseIf Action≟7
              PSE_R := pose_add(PSE_T, p[0,0,0.150,0,0,0])
              PSE_A := pose_add(PSE_T, p[0,0,0.250,0,0,0])
      Case (caseValue=3)
        Folder Output
          'CHANGE THE REFERENCE TO THE FRAME TO MOVE IN'
          Folder define poses
            FRM_Reference := Base
            PSE_T := p[0,0,0,0,0,0]
            PSE_A := pose_add(PSE_T, p[0,0,0.150,0,0,0])
            PSE_R := pose_add(PSE_T, p[0,0,0.100,0,0,0])
      Case (caseValue=5)
        Folder Sarstedt Pickup Table
          'CHANGE THE REFERENCE TO THE FRAME TO MOVE IN'
          Switch expression=JIG
            Case (caseValue=7)
              SuppressedNode
                Folder Sarstedt Rack
                  SuppressedNode
                    Folder Gripping parameters
                      GRP_Open_Pos := 45
                      GRP_Close_Pos := 100
                      Script: rq_set_force_norm(80)
                      Script: rq_set_speed_norm(100)
                  Folder Frame & Position Params
                    Script: FRM_Reference = FRM_SS_SSTable
                    PSE_T := pose_RPY2RotVec(p[0,0,0,0,0,0])
                    PSE_T := pose_trans(PSE_T, GRP_Offset)
                    PSE_A := pose_trans(PSE_T, p[0,0,0.1,0,0,0])
                    PSE_R := pose_add(PSE_T, p[0,0,0.1,0,0,0])
              Folder Sarstedt
                'CHANGE THE REFERENCE TO THE FRAME TO MOVE IN'
                SuppressedNode
                  Folder Gripping parameters
                    GRP_Open_Pos := 45
                    GRP_Close_Pos := 100
                    Script: rq_set_force_norm(80)
                    Script: rq_set_speed_norm(100)
                If TASK.ID≟10
                  Folder Frame & Position Params
                    Script: FRM_Reference = CAM_LM_SSRack
                    PSE_T := uLM_SS_PickPlc
